(* IEC 61131-3 sources: SRCI_CLIENT_PLC/RobotLibrary/Library/POUs/General/MC_RobotTask, 1 file *)

(* ---- MC_RobotTaskFB.st ---- *)
/// Handles multiple mechanisms required for operation of the interface.
/// For maximal performance, this FB must be called after the function FB's,
/// so that the data can be written to the fieldbus in the same cycle as the start of FB occours
FUNCTION_BLOCK MC_RobotTaskFB EXTENDS RobotLibraryLogFB
// -------------------------------------------------------------------------
//  SRCI Robot Library
// -------------------------------------------------------------------------
//
//  Object:      RobotTaskFB
//  Author:      Thorsten Brach
//  Date:        2024-06-01
//
//  Description:
//
//
//  Copyright:
//    (C) 2024 Thorsten Brach. All rights reserved
//             Licensed under the MIT License.
//
//  Disclaimer:
//    This project is provided without any guarantee and can be used for
//    private and commercial purposes. Any use is at the user’s
//    own risk and responsibility.
//
// -------------------------------------------------------------------------
VAR_INPUT
  /// Set TRUE (default) to initialize the interface
  Enable            : BOOL;
  /// User defined robot name
  RobotName         : STRING(20);
  /// Current System Time
  SystemTime        : SystemTime;
  /// Online Change detected
  OnlineChange      : BOOL;
  /// Axes Group ID -> is used to uniquely identify each RA on a per RC basis.
  ///
  /// The IDs start with 0: an RC with only one RA uses ID 0.
  /// ST-FIX F138: spec V1.5.9 says 1 (one RA) and 1-15 (several RAs); this is an error of the spec
  /// (confirmed by PI), the SDK uses 0 too.
  AxesGroupID       : BYTE := 0;
  /// Configuration parameter
  ParCfg            : RobotTaskParCfg;
END_VAR

VAR_IN_OUT
  /// Inputs of PLC for communication from RC
  RobotInData       : ARRAY[*] OF BYTE;
  /// Outputs of PLC for communication to RC
  RobotOutData      : ARRAY[*] OF BYTE;
  ///  User data stored on the PLC according to Table 6-10
  UserData          : UserData;
  /// ToolData stored on PLC. For more information refer to 5.5.6.3
  ToolData          : ARRAY[*] OF Tool;
  /// LoadData stored on PLC.For more information refer to 5.5.6.4
  FrameData         : ARRAY[*] OF Frame;
  /// LoadData stored on PLC.For more information refer to 5.5.6.4
  LoadData          : ARRAY[*] OF Load;
  /// Work areas stored on PLC. For more information refer to 5.5.8
  WorkAreas         : ARRAY[*] OF RobotWorkArea;
  /// Software limits stored on PLC
  SWLimits          : SWLimits;
  /// Default dynamics stored on PLC. For more information refer to 5.5.7
  DefaultDynamics   : DefaultDynamics;
  /// Reference dynamics stored on PLC. For more information refer to 5.5.7
  ReferenceDynamics : ReferenceDynamics;
  /// System log on PLC
  SystemLog         : ARRAY[0..RobotLibraryParameter.SYSTEM_LOG_MAX ] OF STRING(RobotLibraryParameter.MESSAGE_TEXT_LEN);
  /// Message buffer on the PLC - For more information refer to 5.5.11
  MessageLog        : ARRAY[0..RobotLibraryParameter.MESSAGE_LOG_MAX] OF AlarmMessage;
  /// Robot assignment of function
  AxesGroup         : AxesGroup;
END_VAR

VAR_OUTPUT
  /// FB is being processed
  Busy              : BOOL;
  /// Interface is initialized (RI state: "Initialized").
  /// For more information on RI states refer to chapter 5.5.3.1.
  Initialized       : BOOL;
  /// Server and client were successfully synchronized (RI state: "Synchronized").
  /// For more information on the synchronization mechanism refer to chapter 5.6.7.
  Synchronized      : BOOL;
  /// An error occurred
  Error             : BOOL;
  /// ErrorID reported by RC for error identification according to Table 7-1
  ErrorID           : WORD;
  ErrorIdEnum       : RobotLibraryErrorIdEnum;
  ErrorAddTxt       : STRING(RobotLibraryConstants.MAX_ADD_TEXT_LENGTH);
  /// WarningID for warning identification reported during execution of command according to Table 7-3
  WarningID         : WORD;
  WarningIdEnum     : RobotLibraryWarningIdEnum;
  /// InfoID for info identification reported during execution of command according to Table 7-5
  InfoID            : WORD;
  InfoIdEnum        : RobotLibraryInfoIdEnum;
END_VAR

VAR
  /// internal copy of configuration parameter
 _parCfg                       : RobotTaskParCfg;

  /// internal ToolData for comparation to user ToolData
 _toolData                     : ARRAY[0..RobotLibraryParameter.TOOL_MAX       -1] OF Tool;
  /// internal FrameData for comparation to user FrameData
 _frameData                    : ARRAY[0..RobotLibraryParameter.FRAME_MAX      -1] OF Frame;
  /// internal LoadData for comparation to user LoadData
 _loadData                     : ARRAY[0..RobotLibraryParameter.LOAD_MAX       -1] OF Load;
  /// internal WorkAreas for comparation to user WorkAreas
 _workAreas                    : ARRAY[0..RobotLibraryParameter.WORK_AREAS_MAX -1] OF RobotWorkArea;
  /// internal Software limits for comparation to user Software limit
 _swLimits                     : SWLimits;
  /// internal default dynamics for comparation to user default dynamics
 _defaultDynamics              : DefaultDynamics;
  /// internal reference dynamics for comparation to user reference dynamics
 _referenceDynamics            : ReferenceDynamics;

  /// FB for exchange configuration
 _exchangeConfiguration        : MC_ExchangeConfigurationFB;
  /// FB for read robot data
 _readRobotData                : MC_ReadRobotDataFB;
  /// FB for read messaged
 _readMessages                 : MC_ReadMessagesFB;
  /// FB for read tool data
 _readToolData                 : MC_ReadToolDataFB;
  /// FB for read frame data
 _readFrameData                : MC_ReadFrameDataFB;
  /// FB for read load data
 _readLoadData                 : MC_ReadLoadDataFB;
  /// FB for read work area
 _readWorkArea                 : MC_ReadWorkAreaFB;
  /// FB for read robot software limits
 _readRobotSWLimits            : MC_ReadRobotSWLimitsFB;
  /// FB for read robot default dynamics
 _readRobotDefaultDynamics     : MC_ReadRobotDefaultDynamicsFB;
  /// FB for read robot reference dynamics
 _readRobotReferenceDynamics   : MC_ReadRobotReferenceDynamicsFB;

  /// FB for write tool data
 _writeToolData                : MC_WriteToolDataFB;
  /// FB for write frame data
 _writeFrameData               : MC_WriteFrameDataFB;
  /// FB for write load data
 _writeLoadData                : MC_WriteLoadDataFB;
  /// FB for write work area
 _writeWorkArea                : MC_WriteWorkAreaFB;
  /// FB for write robot software limits
 _writeRobotSWLimits           : MC_WriteRobotSWLimitsFB;
  /// FB for write robot default dynamics
 _writeRobotDefaultDynamics    : MC_WriteRobotDefaultDynamicsFB;
  /// FB for write robot reference dynamics
 _writeRobotReferenceDynamics  : MC_WriteRobotReferenceDynamicsFB;
  /// Send Buffer
  SendData                     : RobotLibrarySendDataFB;
  /// Recv Buffer
  RecvData                     : RobotLibraryRecvDataFB;
  /// Telegram
  Telegram                     : Telegram;

  /// internal step counter for command
 _stepCmd                      : DINT;
  /// internal timer for command
  {attribute 'hide'}
 _timerCmd                     : TON;
  /// internal timeout for command
  {attribute 'hide'}
 _timeoutCmd                   : TIME := T#5S;

  /// internal step counter for synchronisation of frame data
 _stepSyncFrameData            : DINT;
  /// internal timer for synchronisation of frame data
  {attribute 'hide'}
 _timerSyncFrameData           : TON;
  /// internal timeout for synchronisation of frame data
  {attribute 'hide'}
 _timeoutSyncFrameData         : TIME := T#5S;
   /// internal index for frame data synchronisation
 _syncIdxFrameData             : USINT;
  /// internal index for maximal amount of frames data( MIN(PLC,RC) )
 _syncIdxMaxFrameData          : DINT;

  /// internal step counter for synchronisation of load data
 _stepSyncLoadData             : DINT;
  /// internal timer for synchronisation of load data
  {attribute 'hide'}
 _timerSyncLoadData             : TON;
  /// internal timeout for synchronisation of load data
  {attribute 'hide'}
 _timeoutSyncLoadData           : TIME := T#5S;
  /// internal index for load data synchronisation
 _syncIdxLoadData               : USINT;
  /// internal index for maximal amount of load data ( MIN(PLC,RC) )
 _syncIdxMaxLoadData            : DINT;

  /// internal step counter for synchronisation of tool data
 _stepSyncToolData              : DINT;
  /// internal timer for synchronisation of tool data
  {attribute 'hide'}
 _timerSyncToolData             : TON;
  /// internal timeout for synchronisation of tool data
  {attribute 'hide'}
 _timeoutSyncToolData           : TIME := T#5S;
  /// internal index for tool data synchronisation
 _syncIdxToolData               : USINT;
  /// internal index for maximal amount of tool data ( MIN(PLC,RC) )
 _syncIdxMaxToolData            : DINT;

  /// internal step counter for synchronisation of work areas
 _stepSyncWorkArea            : DINT;
 /// internal timer for synchronisation of work areas
  {attribute 'hide'}
 _timerSyncWorkArea           : TON;
  /// internal timeout for synchronisation of work areas
  {attribute 'hide'}
 _timeoutSyncWorkArea         : TIME := T#5S;
  /// internal index for WorkArea synchronisation
 _syncIdxWorkArea             : USINT;
  /// internal index for maximal amount of Work Area( MIN(PLC,RC) )
 _syncIdxMaxWorkArea          : DINT;

  /// internal step counter for synchronisation of software limits
 _stepSyncSWLimits            : DINT;
  /// internal timer for synchronisation of software limits
  {attribute 'hide'}
 _timerSyncSWLimits           : TON;
  /// internal timeout for synchronisation of software limits
  {attribute 'hide'}
 _timeoutSyncSWLimits         : TIME := T#5S;

  /// internal step counter for synchronisation of default dynamics
 _stepSyncDefaultDynamics      : DINT;
  /// internal timer for synchronisation of default dynamics
  {attribute 'hide'}
 _timerSyncDefaultDynamics     : TON;
  /// internal timeout for synchronisation of default dynamics
  {attribute 'hide'}
 _timeoutSyncDefaultDynamics   : TIME := T#5S;

  /// internal step counter for synchronisation of reference dynamics
 _stepSyncReferenceDynamics    : DINT;
  /// internal timer for synchronisation of reference dynamics
  {attribute 'hide'}
 _timerSyncReferenceDynamics   : TON;
  /// internal timeout for synchronisation of reference dynamics
  {attribute 'hide'}
 _timeoutSyncReferenceDynamics : TIME := T#5S;

  /// Rising edge for enable
  {attribute 'hide'}
 _enable_R                    : R_TRIG;
  /// Falling edge for enable
  {attribute 'hide'}
 _enable_F                    : F_TRIG;

  /// Flag that indicated the the connection is alive (data exchange)
 _aliveBit                    : BOOL;
  /// last lifesign counter value
 _aliveValue                  : BYTE;
  /// timer for detecting alive state
 _aliveCheck                  : TON;
  /// rising edge for connection is alive
  {attribute 'hide'}
 _alive_R                     : R_TRIG;
  /// falling edge for connection is alive
  {attribute 'hide'}
 _alive_F                     : F_TRIG;
   /// last telegram state
 _lastTelegramState           : TelegramState   := TelegramState.UNDEFINED;
   /// last telegram control
 _lastTelegramControl         : ControlHalfByte := ControlHalfByte.NONE;
END_VAR

VAR // CONSTANT
  /// Lower array dimension of RobotInData
  ROBOT_IN_DATA_MIN   : DINT;
  /// Upper array dimension of RobotInData
  ROBOT_IN_DATA_MAX   : DINT;
  /// Size of RobotInData
  ROBOT_IN_DATA_SIZE  : UDINT;
  /// Lower array dimension of RobotOutData
  ROBOT_OUT_DATA_MIN  : DINT;
  /// Upper array dimension of RobotOutData
  ROBOT_OUT_DATA_MAX  : DINT;
  /// Size of RobotOutData
  ROBOT_OUT_DATA_SIZE : UDINT;
END_VAR

VAR CONSTANT
  {attribute 'hide'}
  FRAGMENT_HEADER_SIZE : UDINT := SIZEOF(TelegramPlcToRobFragmentHeader);
  /// Size of the comand header
  {attribute 'hide'}
  COMMAND_HEADER_SIZE  : UDINT := SIZEOF(TelegramPlcToRobCommandHeader);
  /// Size of the footer
  {attribute 'hide'}
  FOOTER_SIZE          : UDINT := 1;
  /// Minimal payload size for telegram
  {attribute 'hide'}
  MIN_PAYLOAD_SIZE     : UDINT := 1;
  /// Active command
  {attribute 'hide'}
  ACTIVE_CMD           : UDINT := 1;
  /// Buffered command
  {attribute 'hide'}
  BUFFER_CMD           : UDINT := 2;
  /// Empty command entry
  {attribute 'hide'}
  EMPTY_CMD_ENTRY      : AxesGroupAcyclicAcrEntryCmdBuffer := (State := BufferStateCmd.EMPTY);
  /// bitmask to mask the LifeSign out of the halfbyte
  {attribute 'hide'}
  LIFESIGN_BIT_MASK    : BYTE := 2#000_1111;
  /// Primary sequence
  {attribute 'hide'}
  PRIMARY_SEQUENCE     : DINT := 0;
  /// Secondary sequence
  {attribute 'hide'}
  SECONDARY_SEQUENCE   : DINT := 1;
  /// Empty Execution-Order-List entry
  {attribute 'hide'}
  EMPTY_EOL_ENTRY      : DINT := 0;
END_VAR

VAR
  /// ST-FIX F63: telegram sequence that is handled/filled first (lower Seq/Ack number)
  _seqSendFirst : DINT;
  /// ST-FIX F63: loop counter over the telegram sequences in Seq order
  _seqOrderIdx : DINT;
  /// ST-FIX F63: distance of two Seq numbers
  _seqDiff : DINT;
  /// ST-FIX F63: next Seq number
  _seqNext : UINT;
END_VAR

VAR
  /// ST-FIX F65: telegram sequence timeout (4 x LifeSignTimeOut without new Seq number)
  _seqAckTimeout : TON;
  /// ST-FIX F66: lifesign of header and footer differ -> frame is not processed
  _frameInvalid : BOOL;
  /// ST-FIX F79: last error state of the RC during the initialization (reported at the init timeout)
  _initErrorState : TelegramState;
END_VAR

VAR
  _turns : BYTE; // ST-FIX F60: turn number nibble
END_VAR

VAR
  _restartReset : BOOL; // ST-FIX F23: interface reset on the RC requested by a restart
END_VAR

VAR
  /// ST-FIX F132: identification of this instance (1..n, assigned in FB_init, kept by an online change)
 _instanceId : UDINT;
END_VAR

VAR_STAT
  /// ST-FIX F132: number of RobotTask instances created (source of _instanceId)
 _instanceCount   : UDINT;
  /// ST-FIX F132: instance that uses the telegram buffers of the entry (0 = free entry)
 _peripheryOwner  : ARRAY[1..PERIPHERY_ENTRIES] OF UDINT;
  /// ST-FIX F132: address of RobotInData of the entry
 _peripheryInAdr  : ARRAY[1..PERIPHERY_ENTRIES] OF PVOID;
  /// ST-FIX F132: address of RobotOutData of the entry
 _peripheryOutAdr : ARRAY[1..PERIPHERY_ENTRIES] OF PVOID;
END_VAR

VAR CONSTANT
  /// ST-FIX F132: number of RobotTask instances whose telegram buffers are checked
  PERIPHERY_ENTRIES : DINT := 16;
END_VAR

  // Get array dimension of RobotInData
  ROBOT_IN_DATA_MIN  := LOWER_BOUND  ( RobotInData,1);
  ROBOT_IN_DATA_MAX  := UPPER_BOUND  ( RobotInData,1);
  ROBOT_IN_DATA_SIZE := DINT_TO_UDINT( ROBOT_IN_DATA_MAX - ROBOT_IN_DATA_MIN + 1);

  // Get array dimension of RobotInData
  ROBOT_OUT_DATA_MIN  := LOWER_BOUND  ( RobotOutData,1);
  ROBOT_OUT_DATA_MAX  := UPPER_BOUND  ( RobotOutData,1);
  ROBOT_OUT_DATA_SIZE := DINT_TO_UDINT( ROBOT_OUT_DATA_MAX - ROBOT_OUT_DATA_MIN + 1);

  // ST-FIX F132: an AxesGroup and the telegram buffers belong to one RobotTask only (table 7-1:
  // 16#8007 / 16#8008); a second instance does nothing else, so it cannot disturb the first one
  IF ( NOT CheckAssignmentValid( AxesGroup    := AxesGroup,
                                 RobotInData  := RobotInData,
                                 RobotOutData := RobotOutData ) )
  THEN
    Error       := HasError;
    ErrorIdEnum := ErrorID;
    RETURN;
  END_IF

  HandleAxesGroup              ( AxesGroup         := AxesGroup,
  	                             ToolData          := ToolData,
  	                             FrameData         := FrameData,
  	                             LoadData          := LoadData,
  	                             WorkAreas         := WorkAreas,
  	                             SWLimits          := SWLimits,
  	                             DefaultDynamics   := DefaultDynamics,
  	                             ReferenceDynamics := ReferenceDynamics);

  HandleLifeSign               ( AxesGroup         := AxesGroup);
  HandleLogMessagesAck         ( AxesGroup         := AxesGroup);
  HandleInvalidFrames          ( AxesGroup         := AxesGroup, RobotInData := RobotInData);
  HandleTelegramStateCtrl      (                               );
  HandleAliveBit               ( RobotInData[1]                );
  HandleSeqAck                 ( AxesGroup         := AxesGroup);
  HandleUserData               ( AxesGroup         := AxesGroup, UserData := UserData );

  HandleSync                   ( AxesGroup         := AxesGroup,
                                 ToolData          := ToolData,
                                 FrameData         := FrameData,
                                 LoadData          := LoadData,
                                 WorkAreas         := WorkAreas,
                                 SWLimits          := SWLimits,
                                 DefaultDynamics   := DefaultDynamics,
                                 ReferenceDynamics := ReferenceDynamics);

  OnCall                       ( AxesGroup         := AxesGroup);
  OnExecRun                    ( AxesGroup         := AxesGroup);

  AxesGroupToTelegram          ( AxesGroup         := AxesGroup );

  CreateSendPayload            ( AxesGroup         := AxesGroup, RobotOutData := RobotOutData );
  IF ( NOT _frameInvalid ) // ST-FIX F66
  THEN
    ParseRecvPayload             ( AxesGroup         := AxesGroup, RobotInData  := RobotInData);
  END_IF

  AxesGroupFromTelegram        ( AxesGroup         := AxesGroup);

  // call internal functionblocks
  _exchangeConfiguration      ( Name := RobotName, ExecMode := ExecutionMode.PARALLEL, Priority := PriorityLevel.NORMAL, AxesGroup := AxesGroup );
  _readRobotData              ( Name := RobotName, ExecMode := ExecutionMode.PARALLEL, Priority := PriorityLevel.NORMAL, AxesGroup := AxesGroup );
  _readMessages               ( Name := RobotName, ExecMode := ExecutionMode.PARALLEL, Priority := PriorityLevel.NORMAL, AxesGroup := AxesGroup );
  _readToolData               ( UpdateSystemData := FALSE, // ST-FIX F16
   Name := RobotName, ExecMode := ExecutionMode.PARALLEL, Priority := PriorityLevel.NORMAL, AxesGroup := AxesGroup );
  _readFrameData              ( UpdateSystemData := FALSE, // ST-FIX F16
   Name := RobotName, ExecMode := ExecutionMode.PARALLEL, Priority := PriorityLevel.NORMAL, AxesGroup := AxesGroup );
  _readLoadData               ( UpdateSystemData := FALSE, // ST-FIX F16
   Name := RobotName, ExecMode := ExecutionMode.PARALLEL, Priority := PriorityLevel.NORMAL, AxesGroup := AxesGroup );
  _readWorkArea               ( UpdateSystemData := FALSE, // ST-FIX F16
   Name := RobotName, ExecMode := ExecutionMode.PARALLEL, Priority := PriorityLevel.NORMAL, AxesGroup := AxesGroup );
  _readRobotSWLimits          ( UpdateSystemData := FALSE, // ST-FIX F16
   Name := RobotName, ExecMode := ExecutionMode.PARALLEL, Priority := PriorityLevel.NORMAL, AxesGroup := AxesGroup );
  _readRobotDefaultDynamics   ( UpdateSystemData := FALSE, // ST-FIX F16
   Name := RobotName, ExecMode := ExecutionMode.PARALLEL, Priority := PriorityLevel.NORMAL, AxesGroup := AxesGroup );
  _readRobotReferenceDynamics ( UpdateSystemData := FALSE, // ST-FIX F16
   Name := RobotName, ExecMode := ExecutionMode.PARALLEL, Priority := PriorityLevel.NORMAL, AxesGroup := AxesGroup );
  _writeToolData              ( Name := RobotName, ExecMode := ExecutionMode.PARALLEL, Priority := PriorityLevel.NORMAL, AxesGroup := AxesGroup );
  _writeFrameData             ( Name := RobotName, ExecMode := ExecutionMode.PARALLEL, Priority := PriorityLevel.NORMAL, AxesGroup := AxesGroup );
  _writeLoadData              ( Name := RobotName, ExecMode := ExecutionMode.PARALLEL, Priority := PriorityLevel.NORMAL, AxesGroup := AxesGroup );
  _writeWorkArea              ( Name := RobotName, ExecMode := ExecutionMode.PARALLEL, Priority := PriorityLevel.NORMAL, AxesGroup := AxesGroup );
  _writeRobotSWLimits         ( Name := RobotName, ExecMode := ExecutionMode.PARALLEL, Priority := PriorityLevel.NORMAL, AxesGroup := AxesGroup );
  _writeRobotDefaultDynamics  ( Name := RobotName, ExecMode := ExecutionMode.PARALLEL, Priority := PriorityLevel.NORMAL, AxesGroup := AxesGroup );
  _writeRobotReferenceDynamics( Name := RobotName, ExecMode := ExecutionMode.PARALLEL, Priority := PriorityLevel.NORMAL, AxesGroup := AxesGroup );

  // Update SystemLog and MessageLog
  SystemLog  := AxesGroup.MessageLog.SystemLogs;
  MessageLog := AxesGroup.MessageLog.Messages;

END_FUNCTION_BLOCK

METHOD PRIVATE AxesGroupFromTelegram
VAR_IN_OUT
  /// Robot assignment of function
  AxesGroup    : AxesGroup;
END_VAR

  AxesGroupFromTelegramCyclic         (AxesGroup := AxesGroup);
  AxesGroupFromTelegramCyclicOptional (AxesGroup := AxesGroup);

END_METHOD

METHOD PRIVATE AxesGroupFromTelegramCyclic
VAR_IN_OUT
  /// Robot assignment of function
  AxesGroup : AxesGroup;
END_VAR

  // ---------------------------------
  // Mapp Telegramm to AxesGroup Data
  // ---------------------------------
  AxesGroup.Cyclic.RobToPlc.SRCIVersion    := Telegram.RobToPlc.Header.SRCIVersion ;
  AxesGroup.Cyclic.RobToPlc.LifeSign       := Telegram.RobToPlc.Header.LifeSign ;
  AxesGroup.Cyclic.RobToPlc.TelegramState  := Telegram.RobToPlc.Header.TelegramState ;
  AxesGroup.Cyclic.RobToPlc.StatusRobotArm := DwordToRaStatusWord(Telegram.RobToPlc.Header.StatusRobotArm);
  AxesGroup.Cyclic.RobToPlc.Override       := Telegram.RobToPlc.Header.Override ;

END_METHOD

METHOD PRIVATE AxesGroupFromTelegramCyclicOptional
VAR_IN_OUT
  /// Robot assignment of function
  AxesGroup: AxesGroup;
END_VAR

  // Sub ProgramData {{{
  AxesGroup.CyclicOptional.RobToPlc.SubProgramData.Data := Telegram.RobToPlc.CyclicOptional.SubProgramData.Data;
  // }}}

  // Cartesian position {{{
  AxesGroup.CyclicOptional.RobToPlc.CartesianPosition.Active                   :=                                     AxesGroup.CyclicOptional.RobToPlc.CartesianPosition.Active;
  AxesGroup.CyclicOptional.RobToPlc.CartesianPosition.X                        :=                                      Telegram.RobToPlc.CyclicOptional.CartesianPosition.X;
  AxesGroup.CyclicOptional.RobToPlc.CartesianPosition.Y                        :=                                      Telegram.RobToPlc.CyclicOptional.CartesianPosition.Y;
  AxesGroup.CyclicOptional.RobToPlc.CartesianPosition.Z                        :=                                      Telegram.RobToPlc.CyclicOptional.CartesianPosition.Z;
  AxesGroup.CyclicOptional.RobToPlc.CartesianPosition.Rx                       :=                                      Telegram.RobToPlc.CyclicOptional.CartesianPosition.Rx;
  AxesGroup.CyclicOptional.RobToPlc.CartesianPosition.Ry                       :=                                      Telegram.RobToPlc.CyclicOptional.CartesianPosition.Ry;
  AxesGroup.CyclicOptional.RobToPlc.CartesianPosition.Rz                       :=                                      Telegram.RobToPlc.CyclicOptional.CartesianPosition.Rz;
  AxesGroup.CyclicOptional.RobToPlc.CartesianPosition.Config.Shoulder          :=              WordToArmConfigShoulder(Telegram.RobToPlc.CyclicOptional.CartesianPosition.Config);
  AxesGroup.CyclicOptional.RobToPlc.CartesianPosition.Config.Elbow             :=              WordToArmConfigElbow   (Telegram.RobToPlc.CyclicOptional.CartesianPosition.Config);
  AxesGroup.CyclicOptional.RobToPlc.CartesianPosition.Config.Wrist             :=              WordToArmConfigWrist   (Telegram.RobToPlc.CyclicOptional.CartesianPosition.Config);
  _turns := GetHalfeByteLo(Telegram.RobToPlc.CyclicOptional.CartesianPosition.Turns_J2_J1); // ST-FIX F60: sign + magnitude (spec 5.5.4.4)
  AxesGroup.CyclicOptional.RobToPlc.CartesianPosition.TurnNumber.J1Turns := BYTE_TO_SINT(_turns AND 16#07);
  IF ( ( _turns AND 16#08 ) <> 0 )
  THEN
    AxesGroup.CyclicOptional.RobToPlc.CartesianPosition.TurnNumber.J1Turns := INT_TO_SINT(-SINT_TO_INT(AxesGroup.CyclicOptional.RobToPlc.CartesianPosition.TurnNumber.J1Turns));
  END_IF
  _turns := GetHalfeByteHi(Telegram.RobToPlc.CyclicOptional.CartesianPosition.Turns_J2_J1); // ST-FIX F60: sign + magnitude (spec 5.5.4.4)
  AxesGroup.CyclicOptional.RobToPlc.CartesianPosition.TurnNumber.J2Turns := BYTE_TO_SINT(_turns AND 16#07);
  IF ( ( _turns AND 16#08 ) <> 0 )
  THEN
    AxesGroup.CyclicOptional.RobToPlc.CartesianPosition.TurnNumber.J2Turns := INT_TO_SINT(-SINT_TO_INT(AxesGroup.CyclicOptional.RobToPlc.CartesianPosition.TurnNumber.J2Turns));
  END_IF
  _turns := GetHalfeByteLo(Telegram.RobToPlc.CyclicOptional.CartesianPosition.Turns_J4_J3); // ST-FIX F60: sign + magnitude (spec 5.5.4.4)
  AxesGroup.CyclicOptional.RobToPlc.CartesianPosition.TurnNumber.J3Turns := BYTE_TO_SINT(_turns AND 16#07);
  IF ( ( _turns AND 16#08 ) <> 0 )
  THEN
    AxesGroup.CyclicOptional.RobToPlc.CartesianPosition.TurnNumber.J3Turns := INT_TO_SINT(-SINT_TO_INT(AxesGroup.CyclicOptional.RobToPlc.CartesianPosition.TurnNumber.J3Turns));
  END_IF
  _turns := GetHalfeByteHi(Telegram.RobToPlc.CyclicOptional.CartesianPosition.Turns_J4_J3); // ST-FIX F60: sign + magnitude (spec 5.5.4.4)
  AxesGroup.CyclicOptional.RobToPlc.CartesianPosition.TurnNumber.J4Turns := BYTE_TO_SINT(_turns AND 16#07);
  IF ( ( _turns AND 16#08 ) <> 0 )
  THEN
    AxesGroup.CyclicOptional.RobToPlc.CartesianPosition.TurnNumber.J4Turns := INT_TO_SINT(-SINT_TO_INT(AxesGroup.CyclicOptional.RobToPlc.CartesianPosition.TurnNumber.J4Turns));
  END_IF
  _turns := GetHalfeByteLo(Telegram.RobToPlc.CyclicOptional.CartesianPosition.Turns_J6_J5); // ST-FIX F60: sign + magnitude (spec 5.5.4.4)
  AxesGroup.CyclicOptional.RobToPlc.CartesianPosition.TurnNumber.J5Turns := BYTE_TO_SINT(_turns AND 16#07);
  IF ( ( _turns AND 16#08 ) <> 0 )
  THEN
    AxesGroup.CyclicOptional.RobToPlc.CartesianPosition.TurnNumber.J5Turns := INT_TO_SINT(-SINT_TO_INT(AxesGroup.CyclicOptional.RobToPlc.CartesianPosition.TurnNumber.J5Turns));
  END_IF
  _turns := GetHalfeByteHi(Telegram.RobToPlc.CyclicOptional.CartesianPosition.Turns_J6_J5); // ST-FIX F60: sign + magnitude (spec 5.5.4.4)
  AxesGroup.CyclicOptional.RobToPlc.CartesianPosition.TurnNumber.J6Turns := BYTE_TO_SINT(_turns AND 16#07);
  IF ( ( _turns AND 16#08 ) <> 0 )
  THEN
    AxesGroup.CyclicOptional.RobToPlc.CartesianPosition.TurnNumber.J6Turns := INT_TO_SINT(-SINT_TO_INT(AxesGroup.CyclicOptional.RobToPlc.CartesianPosition.TurnNumber.J6Turns));
  END_IF
  AxesGroup.CyclicOptional.RobToPlc.CartesianPosition.TurnNumber.E1Turns := BYTE_TO_SINT(Telegram.RobToPlc.CyclicOptional.CartesianPosition.Turns_E1 AND 16#7F); // ST-FIX F60: sign + magnitude (spec 5.5.4.4)
  IF ( ( Telegram.RobToPlc.CyclicOptional.CartesianPosition.Turns_E1 AND 16#80 ) <> 0 )
  THEN
    AxesGroup.CyclicOptional.RobToPlc.CartesianPosition.TurnNumber.E1Turns := INT_TO_SINT(-SINT_TO_INT(AxesGroup.CyclicOptional.RobToPlc.CartesianPosition.TurnNumber.E1Turns));
  END_IF
  AxesGroup.CyclicOptional.RobToPlc.CartesianPosition.E1                       :=                                      Telegram.RobToPlc.CyclicOptional.CartesianPosition.E1;
  AxesGroup.CyclicOptional.RobToPlc.CartesianPosition.CoordinateSystem.ToolNo  :=                                      Telegram.RobToPlc.CyclicOptional.CartesianPosition.ToolNo; // ST-FIX F59: tool/frame of the returned position
  AxesGroup.CyclicOptional.RobToPlc.CartesianPosition.CurrentCoordinateSystem.ToolNo  :=                                      Telegram.RobToPlc.CyclicOptional.CartesianPosition.CurrentlyUsedToolNo;
  AxesGroup.CyclicOptional.RobToPlc.CartesianPosition.CoordinateSystem.FrameNo :=                                      Telegram.RobToPlc.CyclicOptional.CartesianPosition.FrameNo; // ST-FIX F59: tool/frame of the returned position
  AxesGroup.CyclicOptional.RobToPlc.CartesianPosition.CurrentCoordinateSystem.FrameNo :=                                      Telegram.RobToPlc.CyclicOptional.CartesianPosition.CurrentlyUsedFrameNo;
  // }}}

  // Joint position {{{
  AxesGroup.CyclicOptional.RobToPlc.JointPosition.Active := AxesGroup.CyclicOptional.RobToPlc.JointPosition.Active;
  AxesGroup.CyclicOptional.RobToPlc.JointPosition.J1     :=  Telegram.RobToPlc.CyclicOptional.JointPosition.J1;
  AxesGroup.CyclicOptional.RobToPlc.JointPosition.J2     :=  Telegram.RobToPlc.CyclicOptional.JointPosition.J2;
  AxesGroup.CyclicOptional.RobToPlc.JointPosition.J3     :=  Telegram.RobToPlc.CyclicOptional.JointPosition.J3;
  AxesGroup.CyclicOptional.RobToPlc.JointPosition.J4     :=  Telegram.RobToPlc.CyclicOptional.JointPosition.J4;
  AxesGroup.CyclicOptional.RobToPlc.JointPosition.J5     :=  Telegram.RobToPlc.CyclicOptional.JointPosition.J5;
  AxesGroup.CyclicOptional.RobToPlc.JointPosition.J6     :=  Telegram.RobToPlc.CyclicOptional.JointPosition.J6;
  AxesGroup.CyclicOptional.RobToPlc.JointPosition.E1     :=  Telegram.RobToPlc.CyclicOptional.JointPosition.E1;
  // }}}

  // Force {{{
  AxesGroup.CyclicOptional.RobToPlc.Force.Active          := AxesGroup.CyclicOptional.RobToPlc.Force.Active;
  AxesGroup.CyclicOptional.RobToPlc.Force.X               :=  Telegram.RobToPlc.CyclicOptional.Force.X;
  AxesGroup.CyclicOptional.RobToPlc.Force.Y               :=  Telegram.RobToPlc.CyclicOptional.Force.Y;
  AxesGroup.CyclicOptional.RobToPlc.Force.Z               :=  Telegram.RobToPlc.CyclicOptional.Force.Z;
  AxesGroup.CyclicOptional.RobToPlc.Force.Rx              :=  Telegram.RobToPlc.CyclicOptional.Force.Rx;
  AxesGroup.CyclicOptional.RobToPlc.Force.Ry              :=  Telegram.RobToPlc.CyclicOptional.Force.Ry;
  AxesGroup.CyclicOptional.RobToPlc.Force.Rz              :=  Telegram.RobToPlc.CyclicOptional.Force.Rz;
  // }}}

  // Current {{{
  AxesGroup.CyclicOptional.RobToPlc.Current.Active        := AxesGroup.CyclicOptional.RobToPlc.Current.Active;
  AxesGroup.CyclicOptional.RobToPlc.Current.J1            :=  Telegram.RobToPlc.CyclicOptional.Current.J1;
  AxesGroup.CyclicOptional.RobToPlc.Current.J2            :=  Telegram.RobToPlc.CyclicOptional.Current.J2;
  AxesGroup.CyclicOptional.RobToPlc.Current.J3            :=  Telegram.RobToPlc.CyclicOptional.Current.J3;
  AxesGroup.CyclicOptional.RobToPlc.Current.J4            :=  Telegram.RobToPlc.CyclicOptional.Current.J4;
  AxesGroup.CyclicOptional.RobToPlc.Current.J5            :=  Telegram.RobToPlc.CyclicOptional.Current.J5;
  AxesGroup.CyclicOptional.RobToPlc.Current.J6            :=  Telegram.RobToPlc.CyclicOptional.Current.J6;
  // }}}

  // Two Sequences {{{
  // }}}

  // Cartesian Position Extended
  AxesGroup.CyclicOptional.RobToPlc.CartesianPositionExt.Active := AxesGroup.CyclicOptional.RobToPlc.CartesianPositionExt.Active;
  AxesGroup.CyclicOptional.RobToPlc.CartesianPositionExt.E2     :=  Telegram.RobToPlc.CyclicOptional.CartesianPositionExt.E2;
  AxesGroup.CyclicOptional.RobToPlc.CartesianPositionExt.E3     :=  Telegram.RobToPlc.CyclicOptional.CartesianPositionExt.E3;
  AxesGroup.CyclicOptional.RobToPlc.CartesianPositionExt.E4     :=  Telegram.RobToPlc.CyclicOptional.CartesianPositionExt.E4;
  AxesGroup.CyclicOptional.RobToPlc.CartesianPositionExt.E5     :=  Telegram.RobToPlc.CyclicOptional.CartesianPositionExt.E5;
  AxesGroup.CyclicOptional.RobToPlc.CartesianPositionExt.E6     :=  Telegram.RobToPlc.CyclicOptional.CartesianPositionExt.E6;

  // Joint Position Extended
  AxesGroup.CyclicOptional.RobToPlc.JointPositionExt.Active     := AxesGroup.CyclicOptional.RobToPlc.JointPositionExt.Active;
  AxesGroup.CyclicOptional.RobToPlc.JointPositionExt.E2         :=  Telegram.RobToPlc.CyclicOptional.JointPositionExt.E2;
  AxesGroup.CyclicOptional.RobToPlc.JointPositionExt.E3         :=  Telegram.RobToPlc.CyclicOptional.JointPositionExt.E3;
  AxesGroup.CyclicOptional.RobToPlc.JointPositionExt.E4         :=  Telegram.RobToPlc.CyclicOptional.JointPositionExt.E4;
  AxesGroup.CyclicOptional.RobToPlc.JointPositionExt.E5         :=  Telegram.RobToPlc.CyclicOptional.JointPositionExt.E5;
  AxesGroup.CyclicOptional.RobToPlc.JointPositionExt.E6         :=  Telegram.RobToPlc.CyclicOptional.JointPositionExt.E6;

  // Force Extended
  AxesGroup.CyclicOptional.RobToPlc.ForceExt.Active             := AxesGroup.CyclicOptional.RobToPlc.ForceExt.Active;
  AxesGroup.CyclicOptional.RobToPlc.ForceExt.E1                 :=  Telegram.RobToPlc.CyclicOptional.ForceExt.E1;
  AxesGroup.CyclicOptional.RobToPlc.ForceExt.E2                 :=  Telegram.RobToPlc.CyclicOptional.ForceExt.E2;
  AxesGroup.CyclicOptional.RobToPlc.ForceExt.E3                 :=  Telegram.RobToPlc.CyclicOptional.ForceExt.E3;
  AxesGroup.CyclicOptional.RobToPlc.ForceExt.E4                 :=  Telegram.RobToPlc.CyclicOptional.ForceExt.E4;
  AxesGroup.CyclicOptional.RobToPlc.ForceExt.E5                 :=  Telegram.RobToPlc.CyclicOptional.ForceExt.E5;
  AxesGroup.CyclicOptional.RobToPlc.ForceExt.E6                 :=  Telegram.RobToPlc.CyclicOptional.ForceExt.E6;

  // Current Extended
  AxesGroup.CyclicOptional.RobToPlc.CurrentExt.Active           := AxesGroup.CyclicOptional.RobToPlc.CurrentExt.Active;
  AxesGroup.CyclicOptional.RobToPlc.CurrentExt.E1               :=  Telegram.RobToPlc.CyclicOptional.CurrentExt.E1;
  AxesGroup.CyclicOptional.RobToPlc.CurrentExt.E2               :=  Telegram.RobToPlc.CyclicOptional.CurrentExt.E2;
  AxesGroup.CyclicOptional.RobToPlc.CurrentExt.E3               :=  Telegram.RobToPlc.CyclicOptional.CurrentExt.E3;
  AxesGroup.CyclicOptional.RobToPlc.CurrentExt.E4               :=  Telegram.RobToPlc.CyclicOptional.CurrentExt.E4;
  AxesGroup.CyclicOptional.RobToPlc.CurrentExt.E5               :=  Telegram.RobToPlc.CyclicOptional.CurrentExt.E5;
  AxesGroup.CyclicOptional.RobToPlc.CurrentExt.E6               :=  Telegram.RobToPlc.CyclicOptional.CurrentExt.E6;

END_METHOD

METHOD PRIVATE AxesGroupToTelegram : DINT
VAR_IN_OUT
  /// Robot assignment of function
  AxesGroup : AxesGroup;
END_VAR

VAR
  /// internal index
 _idx                       : DINT;
  /// internal sequence index
 _seqIdx                    : DINT;
  /// internal fragment index
 _fragIdx                   : DINT;
  /// internal register index
 _regIdx                    : DINT;
  /// internal execution order list index
 _listIdx                   : DINT := 1;
  /// internal payload pointer
 _payLoadPtr                : DWORD;
  /// internal fragment action
 _fragmentAction            : FragmentAction;
  /// internal fragment action as string
 _fragmentActionString      : STRING;
  /// maximount amount of bytes per sequence
  SEQUENCE_MAX_PAYLOAD_SIZE : UDINT;
END_VAR

  // ST-FIX F63: the data of a telegram sequence is cleared in AxesGroupToTelegramSequence only
  // when it gets a new Seq number; a sequence that is not acknowledged yet is sent unchanged

  AxesGroupToTelegramHeader        (AxesGroup := AxesGroup);
  AxesGroupToTelegramCyclic        (AxesGroup := AxesGroup);
  AxesGroupToTelegramCyclicOptional(AxesGroup := AxesGroup);
  AxesGroupToTelegramSequence      (AxesGroup := AxesGroup);
  AxesGroupToTelegramFooter        (AxesGroup := AxesGroup);
  AxesGroupToTelegramLogging       (AxesGroup := AxesGroup);

END_METHOD

METHOD PRIVATE AxesGroupToTelegramCyclic : DINT
VAR_IN_OUT
  /// Robot assignment of function
  AxesGroup : AxesGroup;
END_VAR

  IF (AxesGroup.Cyclic.PlcToRob.ToolNo = -1 )
  THEN
    Telegram.PlcToRob.Cyclic.ToolNo  := 16#FF;
  ELSE
    Telegram.PlcToRob.Cyclic.ToolNo  := INT_TO_BYTE(AxesGroup.Cyclic.PlcToRob.ToolNo);
  END_IF

  IF (AxesGroup.Cyclic.PlcToRob.FrameNo = -1 )
  THEN
    Telegram.PlcToRob.Cyclic.FrameNo  := 16#FF;
  ELSE
    Telegram.PlcToRob.Cyclic.FrameNo  := INT_TO_BYTE(AxesGroup.Cyclic.PlcToRob.FrameNo);
  END_IF

END_METHOD

METHOD PRIVATE AxesGroupToTelegramCyclicOptional : DINT
VAR_IN_OUT
  /// Robot assignment of function
  AxesGroup : AxesGroup;
END_VAR

  // AxesGroup.CyclicOptional.PlcToRob.SubProgramData {{{
  IF (AxesGroup.CyclicOptional.PlcToRob.SubProgramData.Active)
  THEN
    Telegram.PlcToRob.CyclicOptional.SubProgramData.Data := AxesGroup.CyclicOptional.PlcToRob.SubProgramData.Data;
  END_IF
  // }}}

  // AxesGroup.CyclicOptional.PlcToRob.CartesianPosition  {{{
  IF (AxesGroup.CyclicOptional.PlcToRob.CartesianPosition.Active)
  THEN
    Telegram.PlcToRob.CyclicOptional.CartesianPosition.X           :=                  AxesGroup.CyclicOptional.PlcToRob.CartesianPosition.X;
    Telegram.PlcToRob.CyclicOptional.CartesianPosition.Y           :=                  AxesGroup.CyclicOptional.PlcToRob.CartesianPosition.Y;
    Telegram.PlcToRob.CyclicOptional.CartesianPosition.Z           :=                  AxesGroup.CyclicOptional.PlcToRob.CartesianPosition.Z;
    Telegram.PlcToRob.CyclicOptional.CartesianPosition.Rx          :=                  AxesGroup.CyclicOptional.PlcToRob.CartesianPosition.Rx;
    Telegram.PlcToRob.CyclicOptional.CartesianPosition.Ry          :=                  AxesGroup.CyclicOptional.PlcToRob.CartesianPosition.Ry;
    Telegram.PlcToRob.CyclicOptional.CartesianPosition.Rz          :=                  AxesGroup.CyclicOptional.PlcToRob.CartesianPosition.Rz;
    Telegram.PlcToRob.CyclicOptional.CartesianPosition.Turns_J2_J1 := CombineHalfSints(AxesGroup.CyclicOptional.PlcToRob.CartesianPosition.TurnNumber.J2Turns,
                                                                                       AxesGroup.CyclicOptional.PlcToRob.CartesianPosition.TurnNumber.J1Turns);
    Telegram.PlcToRob.CyclicOptional.CartesianPosition.Turns_J4_J3 := CombineHalfSints(AxesGroup.CyclicOptional.PlcToRob.CartesianPosition.TurnNumber.J4Turns,
                                                                                       AxesGroup.CyclicOptional.PlcToRob.CartesianPosition.TurnNumber.J3Turns);
    Telegram.PlcToRob.CyclicOptional.CartesianPosition.Turns_J6_J5 := CombineHalfSints(AxesGroup.CyclicOptional.PlcToRob.CartesianPosition.TurnNumber.J6Turns,
                                                                                       AxesGroup.CyclicOptional.PlcToRob.CartesianPosition.TurnNumber.J5Turns);
    // ST-FIX F60: sign + magnitude (spec 5.5.4.4)
    IF ( AxesGroup.CyclicOptional.PlcToRob.CartesianPosition.TurnNumber.E1Turns < 0 )
    THEN
      Telegram.PlcToRob.CyclicOptional.CartesianPosition.Turns_E1 := (INT_TO_BYTE(-SINT_TO_INT(AxesGroup.CyclicOptional.PlcToRob.CartesianPosition.TurnNumber.E1Turns)) AND 16#7F) OR 16#80;
    ELSE
      Telegram.PlcToRob.CyclicOptional.CartesianPosition.Turns_E1 := SINT_TO_BYTE(AxesGroup.CyclicOptional.PlcToRob.CartesianPosition.TurnNumber.E1Turns) AND 16#7F;
    END_IF
  END_IF
  // }}}

  // AxesGroup.CyclicOptional.PlcToRob.CartesianPositionExt {{{
  IF ( AxesGroup.CyclicOptional.PlcToRob.CartesianPositionExt.Active)
  THEN
    Telegram.PlcToRob.CyclicOptional.CartesianPositionExt.E2 := AxesGroup.CyclicOptional.PlcToRob.CartesianPositionExt.E2;
    Telegram.PlcToRob.CyclicOptional.CartesianPositionExt.E3 := AxesGroup.CyclicOptional.PlcToRob.CartesianPositionExt.E3;
    Telegram.PlcToRob.CyclicOptional.CartesianPositionExt.E4 := AxesGroup.CyclicOptional.PlcToRob.CartesianPositionExt.E4;
    Telegram.PlcToRob.CyclicOptional.CartesianPositionExt.E5 := AxesGroup.CyclicOptional.PlcToRob.CartesianPositionExt.E5;
    Telegram.PlcToRob.CyclicOptional.CartesianPositionExt.E6 := AxesGroup.CyclicOptional.PlcToRob.CartesianPositionExt.E6;
  END_IF
  // }}}

  // AxesGroup.CyclicOptional.PlcToRob.JointPosition {{{
  IF ( AxesGroup.CyclicOptional.PlcToRob.JointPosition.Active)
  THEN
    Telegram.PlcToRob.CyclicOptional.JointPosition.J1 := AxesGroup.CyclicOptional.PlcToRob.JointPosition.J1;
    Telegram.PlcToRob.CyclicOptional.JointPosition.J2 := AxesGroup.CyclicOptional.PlcToRob.JointPosition.J2;
    Telegram.PlcToRob.CyclicOptional.JointPosition.J3 := AxesGroup.CyclicOptional.PlcToRob.JointPosition.J3;
    Telegram.PlcToRob.CyclicOptional.JointPosition.J4 := AxesGroup.CyclicOptional.PlcToRob.JointPosition.J4;
    Telegram.PlcToRob.CyclicOptional.JointPosition.J5 := AxesGroup.CyclicOptional.PlcToRob.JointPosition.J5;
    Telegram.PlcToRob.CyclicOptional.JointPosition.J6 := AxesGroup.CyclicOptional.PlcToRob.JointPosition.J6;
    Telegram.PlcToRob.CyclicOptional.JointPosition.E1 := AxesGroup.CyclicOptional.PlcToRob.JointPosition.E1;
  END_IF
  // }}}

  // AxesGroup.CyclicOptional.PlcToRob.JointPositionExt {{{
  IF ( AxesGroup.CyclicOptional.PlcToRob.JointPositionExt.Active)
  THEN
    Telegram.PlcToRob.CyclicOptional.JointPositionExt.E2 := AxesGroup.CyclicOptional.PlcToRob.JointPositionExt.E2;
    Telegram.PlcToRob.CyclicOptional.JointPositionExt.E3 := AxesGroup.CyclicOptional.PlcToRob.JointPositionExt.E3;
    Telegram.PlcToRob.CyclicOptional.JointPositionExt.E4 := AxesGroup.CyclicOptional.PlcToRob.JointPositionExt.E4;
    Telegram.PlcToRob.CyclicOptional.JointPositionExt.E5 := AxesGroup.CyclicOptional.PlcToRob.JointPositionExt.E5;
    Telegram.PlcToRob.CyclicOptional.JointPositionExt.E6 := AxesGroup.CyclicOptional.PlcToRob.JointPositionExt.E6;
  END_IF
  // }}}

  // AxesGroup.CyclicOptional.PlcToRob.Force {{{
  IF ( AxesGroup.CyclicOptional.PlcToRob.Force.Active)
  THEN
    Telegram.PlcToRob.CyclicOptional.Force.X  := AxesGroup.CyclicOptional.PlcToRob.Force.X;
    Telegram.PlcToRob.CyclicOptional.Force.Y  := AxesGroup.CyclicOptional.PlcToRob.Force.Y;
    Telegram.PlcToRob.CyclicOptional.Force.Z  := AxesGroup.CyclicOptional.PlcToRob.Force.Z;
    Telegram.PlcToRob.CyclicOptional.Force.Rx := AxesGroup.CyclicOptional.PlcToRob.Force.Rx;
    Telegram.PlcToRob.CyclicOptional.Force.Ry := AxesGroup.CyclicOptional.PlcToRob.Force.Ry;
    Telegram.PlcToRob.CyclicOptional.Force.Rz := AxesGroup.CyclicOptional.PlcToRob.Force.Rz;
  END_IF
  // }}}

  // AxesGroup.CyclicOptional.PlcToRob.ForceExt {{{
  IF ( AxesGroup.CyclicOptional.PlcToRob.ForceExt.Active)
  THEN
    Telegram.PlcToRob.CyclicOptional.ForceExt.E1 := AxesGroup.CyclicOptional.PlcToRob.ForceExt.E1;
    Telegram.PlcToRob.CyclicOptional.ForceExt.E2 := AxesGroup.CyclicOptional.PlcToRob.ForceExt.E2;
    Telegram.PlcToRob.CyclicOptional.ForceExt.E3 := AxesGroup.CyclicOptional.PlcToRob.ForceExt.E3;
    Telegram.PlcToRob.CyclicOptional.ForceExt.E4 := AxesGroup.CyclicOptional.PlcToRob.ForceExt.E4;
    Telegram.PlcToRob.CyclicOptional.ForceExt.E5 := AxesGroup.CyclicOptional.PlcToRob.ForceExt.E5;
    Telegram.PlcToRob.CyclicOptional.ForceExt.E6 := AxesGroup.CyclicOptional.PlcToRob.ForceExt.E6;
  END_IF
  // }}}

END_METHOD

METHOD PRIVATE AxesGroupToTelegramFooter : DINT
VAR_IN_OUT
  /// Robot assignment of function
  AxesGroup : AxesGroup;
END_VAR

  Telegram.PlcToRob.Footer.LifeSign := GetHalfeByteLo(Telegram.PlcToRob.Header.FastStop_LifeSign);

END_METHOD

METHOD PRIVATE AxesGroupToTelegramHeader : DINT
VAR_IN_OUT
  /// Robot assignment of function
  AxesGroup : AxesGroup;
END_VAR

  Telegram.PlcToRob.Header.SRCIVersion               := VersionToByte(AxesGroup.Cyclic.PlcToRob.SRCIVersion);
  Telegram.PlcToRob.Header.FastStop_LifeSign         := CombineHalfBytes( HalfByteHi := AxesGroup.Cyclic.PlcToRob.FastStop, HalfByteLo := AxesGroup.Cyclic.PlcToRob.LifeSign );
  Telegram.PlcToRob.Header.TelegramLengthPlcToRob    := ParCfg.Com.TelegramLengthPlcToRob;
  Telegram.PlcToRob.Header.TelegramLengthRobToPlc    := ParCfg.Com.TelegramLengthRobToPlc;
  Telegram.PlcToRob.Header.AxesGroupID_Control       := CombineHalfBytes(HalfByteHi := AxesGroup.Cyclic.PlcToRob.AxesGroupID, HalfByteLo := AxesGroup.Cyclic.PlcToRob.Control);
  Telegram.PlcToRob.Header.Reserved                  := 0;
  Telegram.PlcToRob.Header.TelegramNumberPlcToRob    := PlcOptionalCyclicToUint(AxesGroup.Parameter.Plc.OptionalCyclic);
  Telegram.PlcToRob.Header.TelegramNumberRobToPlc    := RobOptionalCyclicToUint(AxesGroup.Parameter.Rob.OptionalCyclic);
  Telegram.PlcToRob.Header.ClientDate                := AxesGroup.Cyclic.PlcToRob.ClientDate;
  Telegram.PlcToRob.Header.ClientTime                := AxesGroup.Cyclic.PlcToRob.ClientTime;

END_METHOD

METHOD PRIVATE AxesGroupToTelegramLogging : DINT
VAR_IN_OUT
  /// Robot assignment of function
  AxesGroup : AxesGroup;
END_VAR

VAR
  /// internal sequence index
 _seqIdx                    : DINT;
  /// internal fragment index
 _fragIdx                   : DINT;
END_VAR

  FOR _seqIdx := 0 TO AxesGroup.State.SequenceCountSend
  DO
    // check new data ?
    IF ( AxesGroup.State.NewSEQ[_seqIdx] )
    THEN
      IF ( Telegram.PlcToRob.Sequence[_seqIdx].Header.PayloadLength > 0 )
      THEN
        // Create log entry
        CreateLogMessagePara4 ( Timestamp   := SystemTime,
                                MessageType := MessageType.CMD,
                                Severity    := Severity.DEBUG,
                                MessageCode := 0,
                                MessageText := 'SendData: SEQ = {1}, added Sequence [{2}] with PayloadLength = {3}, HeaderLength = {4}',
                                Para1       :=  UINT_TO_STRING(Telegram.PlcToRob.Sequence[_seqIdx].Header.SEQ_ACK),
                                Para2       :=  DINT_TO_STRING(_seqIdx),
                                Para3       :=  UINT_TO_STRING(Telegram.PlcToRob.Sequence[_seqIdx].Header.PayloadLength),
                                Para4       :=  DINT_TO_STRING(SIZEOF(Telegram.PlcToRob.Sequence[_seqIdx].Header)));
      END_IF

      FOR _fragIdx := 0 TO AxesGroup.State.FragmentCountSend[_seqIdx]
      DO
        IF ( Telegram.PlcToRob.Sequence[_seqIdx].Fragment[_fragIdx].Header.PayloadLength > 0 )
        THEN
          // Create log entry
          CreateLogMessagePara6 ( Timestamp   := SystemTime,
                                  MessageType := MessageType.CMD,
                                  Severity    := Severity.DEBUG,
                                  MessageCode := 0,
                                  MessageText := 'SendData: added Fragment [{1}] with PayloadLength = {2}, HeaderLength = {3}, CmdID <{4}>, Cmd <{5}> Fragment-Action Bits:{6}' ,
                                  Para1       := DINT_TO_STRING(_fragIdx),
                                  Para2       := UINT_TO_STRING            (Telegram.PlcToRob.Sequence[_seqIdx].Fragment[_fragIdx].Header.PayloadLength),
                                  Para3       := DINT_TO_STRING(SIZEOF     (Telegram.PlcToRob.Sequence[_seqIdx].Fragment[_fragIdx].Header)),
                                  Para4       := UINT_TO_STRING            (Telegram.PlcToRob.Sequence[_seqIdx].Fragment[_fragIdx].Header.CmdID),
                                  Para5       := CMD_TYPE_TO_STRING        (Telegram.PlcToRob.Sequence[_seqIdx].Fragment[_fragIdx].Command.Header.CmdType),
                                  Para6       := FRAGMENT_ACTION_TO_STRING (Telegram.PlcToRob.Sequence[_seqIdx].Fragment[_fragIdx].Header.FragmentAction));

          // Create log entry
          CreateLogMessagePara2 ( Timestamp   := SystemTime,
                                  MessageType := MessageType.CMD,
                                  Severity    := Severity.DEBUG,
                                  MessageCode := 0,
                                  MessageText := 'SendData: added Fragment [{1}] will be executed with ExecMode = [{2}]' ,
                                  Para1       := DINT_TO_STRING(_fragIdx),
                                  Para2       := EXECUTION_MODE_TO_STRING(Telegram.PlcToRob.Sequence[_seqIdx].Fragment[_fragIdx].Command.Header.ExecMode));

        END_IF
      END_FOR
    END_IF
  END_FOR

END_METHOD

METHOD PRIVATE AxesGroupToTelegramSequence : DINT
VAR_IN_OUT
  /// Robot assignment of function
  AxesGroup : AxesGroup;
END_VAR

VAR
  /// internal index
 _idx                       : DINT;
  /// internal sequence index
 _seqIdx                    : DINT;
   /// Amount of sequences
 _seqCount                  : DINT;

  /// internal fragment index
 _fragIdx                   : DINT;
  /// internal register index
 _regIdx                    : DINT;
  /// internal execution order list index
 _listIdx                   : DINT := 1;
  /// internal payload pointer
 _payLoadPtr                : DWORD;
  /// internal fragment action
 _fragmentAction            : FragmentAction;
  /// internal fragment action as string
 _fragmentActionString      : STRING;
  /// maximount amount of bytes per sequence
  SEQUENCE_MAX_PAYLOAD_SIZE : UDINT;

  /// current length of telegram
 _telegramLengthCurrent    : UINT;
END_VAR

  // Check 2nd sequence active ?
  // ST-FIX F67: remaining space for acyclic data at least 1 byte behind the sequence header
  IF ( CalculateSequencePayloadMax(AxesGroup := AxesGroup, Direction := ComDirection.PLC_TO_ROB,
                                   Sequence  := SequenceFlagEnum.PRIMARY_SEQUENCE) < 4 + 1 )
  THEN
    SetError( ErrorID := RobotLibraryErrorIdEnum.ERR_ACYCLIC_AREA_TO_SMALL_PLC_TO_ROB, Overwrite := FALSE );
    // Create log entry
    CreateLogMessage ( Timestamp   := SystemTime,
                       MessageType := MessageType.CMD,
                       Severity    := Severity.ERROR,
                       MessageCode := ErrorID,
                       MessageText := 'Telegram PLC -> RC: no space left for acyclic data');
    RETURN;
  END_IF
  IF ( CalculateSequencePayloadMax(AxesGroup := AxesGroup, Direction := ComDirection.ROB_TO_PLC,
                                   Sequence  := SequenceFlagEnum.PRIMARY_SEQUENCE) < 4 + 1 )
  THEN
    SetError( ErrorID := RobotLibraryErrorIdEnum.ERR_ACYCLIC_AREA_TO_SMALL_ROB_TO_PLC, Overwrite := FALSE );
    // Create log entry
    CreateLogMessage ( Timestamp   := SystemTime,
                       MessageType := MessageType.CMD,
                       Severity    := Severity.ERROR,
                       MessageCode := ErrorID,
                       MessageText := 'Telegram RC -> PLC: no space left for acyclic data');
    RETURN;
  END_IF

  IF ( _parCfg.Com.TwoSequences ) // ST-FIX F63: SEQUENCE_MAX_PAYLOAD_SIZE per sequence, see below
  THEN
    // inc sequence counter
   _seqCount := _seqCount + 1;
  END_IF

  FOR _seqOrderIdx := 0 TO _seqCount
  DO
    // ST-FIX F63: fill the sequence with the lower Seq number first (it is processed first)
    IF ( _seqOrderIdx = 0 )
    THEN
      _seqIdx := _seqSendFirst;
    ELSE
      _seqIdx := 1 - _seqSendFirst;
    END_IF
    // set current SEQ / ACk index
    Telegram.PlcToRob.Sequence[_seqIdx].Header.SEQ_ACK := AxesGroup.State.CurrentSEQ[_seqIdx];

    // only update telegram content if a new sequence SEQ is set
    IF ( AxesGroup.State.NewSEQ[_seqIdx] )
    THEN
      // only reset counters in case of new telegram to send
      // ST-FIX F63: each telegram sequence has its own data area (Fig. 5-205) and starts empty
      IF ( _seqIdx = PRIMARY_SEQUENCE )
      THEN
        SEQUENCE_MAX_PAYLOAD_SIZE := CalculateSequencePayloadMax(AxesGroup := AxesGroup,
                                                                 Direction := ComDirection.PLC_TO_ROB,
                                                                 Sequence  := SequenceFlagEnum.PRIMARY_SEQUENCE);
      ELSE
        SEQUENCE_MAX_PAYLOAD_SIZE := CalculateSequencePayloadMax(AxesGroup := AxesGroup,
                                                                 Direction := ComDirection.PLC_TO_ROB,
                                                                 Sequence  := SequenceFlagEnum.SECONDARY_SEQUENCE);
      END_IF
      Telegram.PlcToRob.Sequence[_seqIdx].Header.PayloadLength := 0;
      FOR _idx := 0 TO RobotLibraryParameter.FRAGMENT_MAX
      DO
        Telegram.PlcToRob.Sequence[_seqIdx].Fragment[_idx].Header.PayloadLength := 0;
      END_FOR
     _fragIdx := 0;
     _listIdx := 1;
      AxesGroup.State.FragmentCountSend[_seqIdx] := 0;

      // calc current telegram payload length
     _telegramLengthCurrent := 4 + Telegram.PlcToRob.Sequence[_seqIdx].Header.PayloadLength; // ST-FIX F63: sequence header + payload

      // Bedingung anpassen und TWO_SEQUENCES berücksichtigen
      WHILE ( _telegramLengthCurrent + FRAGMENT_HEADER_SIZE + MIN_PAYLOAD_SIZE <= SEQUENCE_MAX_PAYLOAD_SIZE ) // ST-FIX F63
      DO
        // Check command in Execution-Order-List available ?
        IF ( AxesGroup.Acyclic.ActiveCommandRegister.ExecutionOrderList[_listIdx] > EMPTY_EOL_ENTRY)
        THEN
          // set current SEQ / ACk index
          Telegram.PlcToRob.Sequence[_seqIdx].Header.SEQ_ACK := AxesGroup.State.CurrentSEQ[_seqIdx];

          // get active command register index
         _regIdx := AxesGroup.Acyclic.ActiveCommandRegister.ExecutionOrderList[_listIdx];

          // check State of the current ACR entry ?
          IF (( AxesGroup.Acyclic.ActiveCommandRegister.Register[_regIdx].Command[ACTIVE_CMD].State >= BufferStateCmd.CREATED  ) AND
              ( AxesGroup.Acyclic.ActiveCommandRegister.Register[_regIdx].Command[ACTIVE_CMD].State <= BufferStateCmd.SENDING  ))
          THEN
            // add size of fragement header
            Telegram.PlcToRob.Sequence[_seqIdx].Header.PayloadLength :=
              Telegram.PlcToRob.Sequence[_seqIdx].Header.PayloadLength + SIZEOF(Telegram.PlcToRob.Sequence[_seqIdx].Fragment[_fragIdx].Header);

            Telegram.PlcToRob.Sequence[_seqIdx].Fragment[_fragIdx].Header.CmdID          := AxesGroup.Acyclic.ActiveCommandRegister.Register[_regIdx].UniqueID;
            Telegram.PlcToRob.Sequence[_seqIdx].Fragment[_fragIdx].Header.Reserve        := 0;
            Telegram.PlcToRob.Sequence[_seqIdx].Fragment[_fragIdx].Header.FragmentAction := 0; // will be set below
            Telegram.PlcToRob.Sequence[_seqIdx].Fragment[_fragIdx].Header.PayloadPointer := AxesGroup.Acyclic.ActiveCommandRegister.Register[_regIdx].Command[ACTIVE_CMD].PayLoadPtr;

            // The 1st message resets the ACR entry on the server side
           _fragmentAction.Reset := (( AxesGroup.Acyclic.ActiveCommandRegister.Register[_regIdx].Command[ACTIVE_CMD].State      = BufferStateCmd.CREATED ) AND
                                     ( AxesGroup.Acyclic.ActiveCommandRegister.Register[_regIdx].Command[ACTIVE_CMD].PayLoadPtr = 0                      ));

            // Update messages must clear the ACR entry on the server side
           _fragmentAction.Clear := (( AxesGroup.Acyclic.ActiveCommandRegister.Register[_regIdx].Command[ACTIVE_CMD].State      = BufferStateCmd.UPDATE_AVAILABLE  ) AND
                                     ( AxesGroup.Acyclic.ActiveCommandRegister.Register[_regIdx].Command[ACTIVE_CMD].PayLoadPtr = 0                                ));

            // fill telegramm header - just for later debugging ( the header is part of the command payload itselfy ) {{{
            Telegram.PlcToRob.Sequence[_seqIdx].Fragment[_fragIdx].Command.Header.CmdType       := CombineBytesToUint ( AxesGroup.Acyclic.ActiveCommandRegister.Register[_regIdx].Command[ACTIVE_CMD].Payload[0],
                                                                                                                        AxesGroup.Acyclic.ActiveCommandRegister.Register[_regIdx].Command[ACTIVE_CMD].Payload[1]);
            Telegram.PlcToRob.Sequence[_seqIdx].Fragment[_fragIdx].Command.Header.ExecMode.0    :=                      AxesGroup.Acyclic.ActiveCommandRegister.Register[_regIdx].Command[ACTIVE_CMD].Payload[2].0;
            Telegram.PlcToRob.Sequence[_seqIdx].Fragment[_fragIdx].Command.Header.ExecMode.1    :=                      AxesGroup.Acyclic.ActiveCommandRegister.Register[_regIdx].Command[ACTIVE_CMD].Payload[2].1;
            Telegram.PlcToRob.Sequence[_seqIdx].Fragment[_fragIdx].Command.Header.ExecMode.2    :=                      AxesGroup.Acyclic.ActiveCommandRegister.Register[_regIdx].Command[ACTIVE_CMD].Payload[2].2;
            Telegram.PlcToRob.Sequence[_seqIdx].Fragment[_fragIdx].Command.Header.ExecMode.3    :=                      AxesGroup.Acyclic.ActiveCommandRegister.Register[_regIdx].Command[ACTIVE_CMD].Payload[2].3;
            Telegram.PlcToRob.Sequence[_seqIdx].Fragment[_fragIdx].Command.Header.Prio.0        :=                      AxesGroup.Acyclic.ActiveCommandRegister.Register[_regIdx].Command[ACTIVE_CMD].Payload[3].0;
            Telegram.PlcToRob.Sequence[_seqIdx].Fragment[_fragIdx].Command.Header.Prio.1        :=                      AxesGroup.Acyclic.ActiveCommandRegister.Register[_regIdx].Command[ACTIVE_CMD].Payload[3].1;
            Telegram.PlcToRob.Sequence[_seqIdx].Fragment[_fragIdx].Command.Header.Prio.2        :=                      AxesGroup.Acyclic.ActiveCommandRegister.Register[_regIdx].Command[ACTIVE_CMD].Payload[3].2;
            Telegram.PlcToRob.Sequence[_seqIdx].Fragment[_fragIdx].Command.Header.Prio.3        :=                      AxesGroup.Acyclic.ActiveCommandRegister.Register[_regIdx].Command[ACTIVE_CMD].Payload[3].3;
            Telegram.PlcToRob.Sequence[_seqIdx].Fragment[_fragIdx].Command.Header.ParSequence.0 :=                      AxesGroup.Acyclic.ActiveCommandRegister.Register[_regIdx].Command[ACTIVE_CMD].Payload[3].4;
            Telegram.PlcToRob.Sequence[_seqIdx].Fragment[_fragIdx].Command.Header.ParSequence.1 :=                      AxesGroup.Acyclic.ActiveCommandRegister.Register[_regIdx].Command[ACTIVE_CMD].Payload[3].5;
            Telegram.PlcToRob.Sequence[_seqIdx].Fragment[_fragIdx].Command.Header.ParSequence.2 :=                      AxesGroup.Acyclic.ActiveCommandRegister.Register[_regIdx].Command[ACTIVE_CMD].Payload[3].6;
            Telegram.PlcToRob.Sequence[_seqIdx].Fragment[_fragIdx].Command.Header.ParSequence.3 :=                      AxesGroup.Acyclic.ActiveCommandRegister.Register[_regIdx].Command[ACTIVE_CMD].Payload[3].7;
            // }}}
            // loop through the payload
            FOR _payLoadPtr := AxesGroup.Acyclic.ActiveCommandRegister.Register[_regIdx].Command[ACTIVE_CMD].PayLoadPtr TO AxesGroup.Acyclic.ActiveCommandRegister.Register[_regIdx].Command[ACTIVE_CMD].PayloadLen -1
            DO
              // copy payload
              Telegram.PlcToRob.Sequence[_seqIdx].Fragment[_fragIdx].Command.Payload[_payLoadPtr]
                := AxesGroup.Acyclic.ActiveCommandRegister.Register[_regIdx].Command[ACTIVE_CMD].Payload[_payLoadPtr];

              // inc current sequence payload length
              Telegram.PlcToRob.Sequence[_seqIdx].Header.PayloadLength
                := Telegram.PlcToRob.Sequence[_seqIdx].Header.PayloadLength + 1;

              // inc current fragment payload length
              Telegram.PlcToRob.Sequence[_seqIdx].Fragment[_fragIdx].Header.PayloadLength
                := Telegram.PlcToRob.Sequence[_seqIdx].Fragment[_fragIdx].Header.PayloadLength + 1;

              // inc payload pointer in active command register
              AxesGroup.Acyclic.ActiveCommandRegister.Register[_regIdx].Command[ACTIVE_CMD].PayLoadPtr
                := AxesGroup.Acyclic.ActiveCommandRegister.Register[_regIdx].Command[ACTIVE_CMD].PayLoadPtr + 1;

              // set command state
              IF ( AxesGroup.Acyclic.ActiveCommandRegister.Register[_regIdx].Command[ACTIVE_CMD].PayLoadPtr >= AxesGroup.Acyclic.ActiveCommandRegister.Register[_regIdx].Command[ACTIVE_CMD].PayLoadLen)
              THEN
                AxesGroup.Acyclic.ActiveCommandRegister.Register[_regIdx].Command[ACTIVE_CMD].State := BufferStateCmd.PROCESSED;
              ELSE
                AxesGroup.Acyclic.ActiveCommandRegister.Register[_regIdx].Command[ACTIVE_CMD].State := BufferStateCmd.SENDING;
              END_IF

              // calc current telegram payload length
             _telegramLengthCurrent := 4 + Telegram.PlcToRob.Sequence[_seqIdx].Header.PayloadLength; // ST-FIX F63: sequence header + payload

              // check limit reached ?
              IF ( _telegramLengthCurrent >= SEQUENCE_MAX_PAYLOAD_SIZE (* ST-FIX F63 *))
              THEN
                EXIT; // -> abort for loop
              END_IF
            END_FOR

            // check payload complete ?
           _fragmentAction.Complete := AxesGroup.Acyclic.ActiveCommandRegister.Register[_regIdx].Command[ACTIVE_CMD].PayLoadPtr
                                    >= AxesGroup.Acyclic.ActiveCommandRegister.Register[_regIdx].Command[ACTIVE_CMD].PayloadLen;

            // just for brakepoint
            IF (_fragmentAction.Complete)
            THEN
             _fragmentAction.Complete := _fragmentAction.Complete;
            END_IF

            // set fragment action
            Telegram.PlcToRob.Sequence[_seqIdx].Fragment[_fragIdx].Header.FragmentAction := FragmentActionToByte(_fragmentAction);
          END_IF
        END_IF

        // inc execution order list index
       _listIdx := _listIdx + 1;
        // inc fragment index
       _fragIdx := _fragIdx + 1;

        // check abort conditions
        IF (( _telegramLengthCurrent                                                >= SEQUENCE_MAX_PAYLOAD_SIZE (* ST-FIX F63 *)  ) OR  // Payload limit reached
            ( _fragIdx                                                              >=  RobotLibraryParameter.FRAGMENT_MAX ) OR  // Max fragment limit reached
            (  AxesGroup.Acyclic.ActiveCommandRegister.ExecutionOrderList[_listIdx]  =  EMPTY_EOL_ENTRY                    ))    // No entry in ExecutionOrderList left
        THEN
          EXIT;// -> Abort while loop
        END_IF
      END_WHILE

      AxesGroup.State.SequenceCountSend          := _seqCount; // ST-FIX F63
      AxesGroup.State.FragmentCountSend[_seqIdx] := _fragIdx;

    END_IF
  END_FOR

END_METHOD

METHOD CalculateCyclicDataLength : UINT
VAR_IN_OUT
  /// Robot assignment of function
  AxesGroup : AxesGroup;
END_VAR
VAR_INPUT
  /// Communication direction
  Direction : ComDirection;
END_VAR

VAR CONSTANT
  /// Size of the header
  ROB_TO_PLC_HEADER_SIZE : UINT := 10;
END_VAR

  // ------------------------------------
  // PLC -> ROB
  // ------------------------------------
  IF (Direction = ComDirection.PLC_TO_ROB)
  THEN
    // Add Header size
    CalculateCyclicDataLength := CalculateCyclicDataLength + SIZEOF(Telegram.PlcToRob.Header);
    // Add Cyclic size (ST-FIX F2: only with Cartesian Position RC -> PLC)
    IF ( AxesGroup.CyclicOptional.RobToPlc.CartesianPosition.Active )
    THEN
      CalculateCyclicDataLength := CalculateCyclicDataLength + SIZEOF(Telegram.PlcToRob.Cyclic);
    END_IF

    // Check SubProgramData active ?
    IF ( AxesGroup.CyclicOptional.PlcToRob.SubProgramData.Active )
    THEN
      // Add SubProgramData size
      CalculateCyclicDataLength := CalculateCyclicDataLength + SIZEOF(Telegram.PlcToRob.CyclicOptional.SubProgramData);
    END_IF

    // Check CartesianPosition active ?
    IF ( AxesGroup.CyclicOptional.PlcToRob.CartesianPosition.Active )
    THEN
      // Add CartesianPosition size
      CalculateCyclicDataLength := CalculateCyclicDataLength + SIZEOF(Telegram.PlcToRob.CyclicOptional.CartesianPosition);
    END_IF

    // Check JointPosition active ?
    IF ( AxesGroup.CyclicOptional.PlcToRob.JointPosition.Active )
    THEN
      // Add JointPosition size
      CalculateCyclicDataLength := CalculateCyclicDataLength + SIZEOF(Telegram.PlcToRob.CyclicOptional.JointPosition);
    END_IF

    // Check Force active ?
    IF ( AxesGroup.CyclicOptional.PlcToRob.Force.Active )
    THEN
      // Add Force size
      CalculateCyclicDataLength := CalculateCyclicDataLength + SIZEOF(Telegram.PlcToRob.CyclicOptional.Force);
    END_IF

    // Check CartesianPositionExt acive ?
    IF ( AxesGroup.CyclicOptional.PlcToRob.CartesianPositionExt.Active )
    THEN
      // Add CartesianPositionExt size
      CalculateCyclicDataLength := CalculateCyclicDataLength + SIZEOF(Telegram.PlcToRob.CyclicOptional.CartesianPositionExt);
    END_IF

    // Check JointPositionExt active ?
    IF ( AxesGroup.CyclicOptional.PlcToRob.JointPositionExt.Active )
    THEN
      // Add JointPositionExt size
      CalculateCyclicDataLength := CalculateCyclicDataLength + SIZEOF(Telegram.PlcToRob.CyclicOptional.JointPositionExt);
    END_IF

    // Check ForceExt active ?
    IF ( AxesGroup.CyclicOptional.PlcToRob.ForceExt.Active )
    THEN
      // Add ForceExt size
      CalculateCyclicDataLength := CalculateCyclicDataLength + SIZEOF(Telegram.PlcToRob.CyclicOptional.ForceExt);
    END_IF
  END_IF

  // ------------------------------------
  // ROB -> PLC
  // ------------------------------------
  IF (Direction = ComDirection.ROB_TO_PLC)
  THEN
    // Add Header size
    CalculateCyclicDataLength := CalculateCyclicDataLength + ROB_TO_PLC_HEADER_SIZE;
    // a constant, because SIZEOF(Telegram.RobToPlc.Header) counts the VersionStruct instead of one byte

    // Check SubProgramData active ?
    IF ( AxesGroup.CyclicOptional.RobToPlc.SubProgramData.Active )
    THEN
      // Add SubProgramData size
      CalculateCyclicDataLength := CalculateCyclicDataLength + SIZEOF(Telegram.RobToPlc.CyclicOptional.SubProgramData);
    END_IF

    // Check CartesianPosition active ?
    IF ( AxesGroup.CyclicOptional.RobToPlc.CartesianPosition.Active )
    THEN
      // Add CartesianPosition size
      CalculateCyclicDataLength := CalculateCyclicDataLength + SIZEOF(Telegram.RobToPlc.CyclicOptional.CartesianPosition);
    END_IF

    // Check JointPosition active ?
    IF ( AxesGroup.CyclicOptional.RobToPlc.JointPosition.Active )
    THEN
      // Add JointPosition size
      CalculateCyclicDataLength := CalculateCyclicDataLength + SIZEOF(Telegram.RobToPlc.CyclicOptional.JointPosition);
    END_IF

    // Check Force active ?
    IF ( AxesGroup.CyclicOptional.RobToPlc.Force.Active )
    THEN
      // Add Force size
      CalculateCyclicDataLength := CalculateCyclicDataLength + SIZEOF(Telegram.RobToPlc.CyclicOptional.Force);
    END_IF

    // Check Current acive ?
    IF ( AxesGroup.CyclicOptional.RobToPlc.Current.Active )
    THEN
      // Add Current size
      CalculateCyclicDataLength := CalculateCyclicDataLength + SIZEOF(Telegram.RobToPlc.CyclicOptional.Current);
    END_IF

    // Check CartesianPositionExt acive ?
    IF ( AxesGroup.CyclicOptional.RobToPlc.CartesianPositionExt.Active )
    THEN
      // Add CartesianPositionExt size
      CalculateCyclicDataLength := CalculateCyclicDataLength + SIZEOF(Telegram.RobToPlc.CyclicOptional.CartesianPositionExt);
    END_IF

    // Check JointPositionExt active ?
    IF ( AxesGroup.CyclicOptional.RobToPlc.JointPositionExt.Active )
    THEN
      // Add JointPositionExt size
      CalculateCyclicDataLength := CalculateCyclicDataLength + SIZEOF(Telegram.RobToPlc.CyclicOptional.JointPositionExt);
    END_IF

    // Check ForceExt active ?
    IF ( AxesGroup.CyclicOptional.RobToPlc.ForceExt.Active )
    THEN
      // Add ForceExt size
      CalculateCyclicDataLength := CalculateCyclicDataLength + SIZEOF(Telegram.RobToPlc.CyclicOptional.ForceExt);
    END_IF

    // Check CurrentExt active ?
    IF ( AxesGroup.CyclicOptional.RobToPlc.CurrentExt.Active )
    THEN
      // Add CurrentExt size
      CalculateCyclicDataLength := CalculateCyclicDataLength + SIZEOF(Telegram.RobToPlc.CyclicOptional.CurrentExt);
    END_IF
  END_IF

END_METHOD

METHOD CalculateSequencePayloadMax : UINT
VAR_IN_OUT
  /// Robot assignment of function
  AxesGroup : AxesGroup;
END_VAR
VAR_INPUT
  /// Communication direction
  Direction : ComDirection;
  /// Sequeunce
  Sequence : SequenceFlag;
END_VAR

VAR
  /// Length of the cyclic header
 _cyclicDataLength      : UINT;
  /// Acyclic area (ST-FIX F63)
 _area                  : UDINT;
END_VAR

  // calculate cyclic header length
  _cyclicDataLength := CalculateCyclicDataLength(AxesGroup := AxesGroup, Direction := Direction);

  // ST-FIX F63: acyclic area without the footer, halved for two sequences (spec Fig. 5-205)
  IF ( Direction = ComDirection.PLC_TO_ROB )
  THEN
    _area := UINT_TO_UDINT(_parCfg.Com.TelegramLengthPlcToRob) - UINT_TO_UDINT(_cyclicDataLength) - FOOTER_SIZE;
  ELSE
    _area := UINT_TO_UDINT(_parCfg.Com.TelegramLengthRobToPlc) - UINT_TO_UDINT(_cyclicDataLength) - FOOTER_SIZE;
  END_IF

  IF ( NOT _parCfg.Com.TwoSequences )
  THEN
    IF ( Sequence = SequenceFlag.PRIMARY_SEQUENCE )
    THEN
      CalculateSequencePayloadMax := UDINT_TO_UINT(_area);
    ELSE
      CalculateSequencePayloadMax := 0;
    END_IF
  ELSIF ( Sequence = SequenceFlag.PRIMARY_SEQUENCE )
  THEN
    CalculateSequencePayloadMax := UDINT_TO_UINT(_area / 2);
  ELSE
    CalculateSequencePayloadMax := UDINT_TO_UINT(_area - _area / 2);
  END_IF

END_METHOD

METHOD CalculateSequencePayloadStartAdr : UINT
VAR_IN_OUT
  /// Robot assignment of function
  AxesGroup : AxesGroup;
END_VAR
VAR_INPUT
  /// Communication direction
  Direction : ComDirection;
  /// Sequeunce
  Sequence : SequenceFlag;
END_VAR

VAR
  /// Length of the cyclic header
 _cyclicDataLength      : UINT;
  /// Length of the sequnce payload
 _sequencePayloadLength : UINT;
END_VAR

  // calculate cyclic header length
  _cyclicDataLength := CalculateCyclicDataLength(AxesGroup := AxesGroup, Direction := Direction);

  CASE (Sequence)
  OF

    SequenceFlag.PRIMARY_SEQUENCE   :

      // return start address
      CalculateSequencePayloadStartAdr := _cyclicDataLength;

    SequenceFlag.SECONDARY_SEQUENCE :

      // calculate sequence payload max
     _sequencePayloadLength
       := CalculateSequencePayloadMax( AxesGroup := AxesGroup,
                                       Direction := Direction,
                                       Sequence  := SequenceFlag.PRIMARY_SEQUENCE ); // ST-FIX F63: behind the area of the 1st sequence

      // return start address
      CalculateSequencePayloadStartAdr := _cyclicDataLength + _sequencePayloadLength;

  END_CASE

END_METHOD

METHOD PROTECTED CalculateTelegramLengthPlcToRob : UINT
VAR_IN_OUT
  /// Robot assignment of function
  AxesGroup : AxesGroup;
END_VAR
VAR
  /// length of the cyclic data block
 _cyclicDataLength : UINT;
END_VAR

  _cyclicDataLength := CalculateCyclicDataLength(AxesGroup := AxesGroup, Direction := ComDirection.PLC_TO_ROB);

  IF ( _parCfg.Com.TwoSequences )
  THEN
    CalculateTelegramLengthPlcToRob := _cyclicDataLength
                                      + SIZEOF(Telegram.PlcToRob.Sequence[  PRIMARY_SEQUENCE].Header)
                                      +       (Telegram.PlcToRob.Sequence[  PRIMARY_SEQUENCE].Header.PayloadLength)
                                      + SIZEOF(Telegram.PlcToRob.Sequence[SECONDARY_SEQUENCE].Header)
                                      +       (Telegram.PlcToRob.Sequence[SECONDARY_SEQUENCE].Header.PayloadLength)
                                      + SIZEOF(Telegram.PlcToRob.Footer);
  ELSE
    CalculateTelegramLengthPlcToRob := _cyclicDataLength
                                      + SIZEOF(Telegram.PlcToRob.Sequence[PRIMARY_SEQUENCE].Header)
                                      +       (Telegram.PlcToRob.Sequence[PRIMARY_SEQUENCE].Header.PayloadLength)
                                      + SIZEOF(Telegram.PlcToRob.Footer);
  END_IF

END_METHOD

/// ST-FIX F132: checks that the AxesGroup and the telegram buffers are not used by another RobotTask
/// (table 7-1: 16#8007 ERR_AXESGROUP_INVALID, 16#8008 ERR_PERIPHERY_INVALID) and registers them
METHOD PRIVATE CheckAssignmentValid : BOOL
VAR_IN_OUT
  /// Robot assignment of function
  AxesGroup    : AxesGroup;
  /// Inputs of PLC for communication from RC
  RobotInData  : ARRAY[*] OF BYTE;
  /// Outputs of PLC for communication to RC
  RobotOutData : ARRAY[*] OF BYTE;
END_VAR
VAR
  /// Loop index over the entries
 _idx     : DINT;
  /// Entry of this instance
 _own     : DINT;
  /// First free entry
 _free    : DINT;
  /// Address of RobotInData
 _inAdr   : PVOID;
  /// Address of RobotOutData
 _outAdr  : PVOID;
END_VAR

  CheckAssignmentValid := FALSE;

  // AxesGroup used by another RobotTask ?
  IF (( AxesGroup.State.RobotTaskId <> 0           ) AND
      ( AxesGroup.State.RobotTaskId <> _instanceId ))
  THEN
    IF ( ErrorID <> RobotLibraryErrorIdEnum.ERR_AXESGROUP_INVALID )
    THEN
      SetError( ErrorID := RobotLibraryErrorIdEnum.ERR_AXESGROUP_INVALID, Overwrite := TRUE );
      // Create log entry
      CreateLogMessagePara1 ( Timestamp   := SystemTime,
                              MessageType := MessageType.CMD,
                              Severity    := Severity.ERROR,
                              MessageCode := ErrorID,
                              MessageText := 'AxesGroup is already used by RobotTask {1}',
                              Para1       := UDINT_TO_STRING(AxesGroup.State.RobotTaskId));
    END_IF
    RETURN;
  END_IF

  // telegram buffers used by another RobotTask ?
  _inAdr  := ADR(RobotInData [ROBOT_IN_DATA_MIN ]);
  _outAdr := ADR(RobotOutData[ROBOT_OUT_DATA_MIN]);
  _own    := 0;
  _free   := 0;
  FOR _idx := 1 TO PERIPHERY_ENTRIES
  DO
    IF ( _peripheryOwner[_idx] = _instanceId )
    THEN
     _own := _idx;
    ELSIF ( _peripheryOwner[_idx] = 0 )
    THEN
      IF ( _free = 0 )
      THEN
       _free := _idx;
      END_IF
    ELSIF (( _peripheryInAdr [_idx] = _inAdr  ) OR
           ( _peripheryOutAdr[_idx] = _outAdr ))
    THEN
      IF ( ErrorID <> RobotLibraryErrorIdEnum.ERR_PERIPHERY_INVALID )
      THEN
        SetError( ErrorID := RobotLibraryErrorIdEnum.ERR_PERIPHERY_INVALID, Overwrite := TRUE );
        // Create log entry
        CreateLogMessagePara1 ( Timestamp   := SystemTime,
                                MessageType := MessageType.CMD,
                                Severity    := Severity.ERROR,
                                MessageCode := ErrorID,
                                MessageText := 'Telegram buffers are already used by RobotTask {1}',
                                Para1       := UDINT_TO_STRING(_peripheryOwner[_idx]));
      END_IF
      RETURN;
    END_IF
  END_FOR

  // register this instance (the addresses can change after an online change)
  IF ( _own = 0 )
  THEN
   _own := _free;
  END_IF
  IF ( _own > 0 )
  THEN
   _peripheryOwner [_own] := _instanceId;
   _peripheryInAdr [_own] := _inAdr;
   _peripheryOutAdr[_own] := _outAdr;
  END_IF
  AxesGroup.State.RobotTaskId := _instanceId;

  CheckAssignmentValid := TRUE;

END_METHOD

METHOD PROTECTED CheckParameterChanged : BOOL
VAR_IN_OUT
  /// Robot assignment of function
  AxesGroup    : AxesGroup;
END_VAR

VAR
  /// internal index for loops
 _idx : DINT;
END_VAR

  // Check initialization is already done ?
  IF ( NOT Initialized )
  THEN
    CheckParameterChanged := FALSE;
    RETURN;
  END_IF

  // compare memory
  CheckParameterChanged := ( SysDepMemCmp(pData1 := ADR(ParCfg), pData2 := ADR(_parCfg), DataLen := SIZEOF(ParCfg)) <> RobotLibraryConstants.OK );

  FOR _idx := SyncTime.DURING_START_UP TO SyncTime.AFTER_START_UP
  DO
    // Check Tool SyncMode changed ?
    IF ( _parCfg.Plc.Parameter.SynchronizationModes.Tool[_idx] <> ParCfg.Plc.Parameter.SynchronizationModes.Tool[_idx] )
    THEN
      // Set info
      SetInfo( InfoID := RobotLibraryInfoIdEnum.INFO_CHANGE_TOOL_SYNC_MODE_TO_NEGATIVE_ONLY_AT_PLC_START_ALLOWED, Overwrite := TRUE);

      // Create log entry
      CreateLogMessagePara3( Timestamp   := SystemTime,
                             MessageType := MessageType.CMD,
                             Severity    := Severity.INFO,
                             MessageCode := 0,
                             MessageText := 'SyncMode.Tool[{1}] changed from {2} to {3}, but this is only allowed at PLC start',
                             Para1       := SYNC_TIME_TO_STRING(_idx),
                             Para2       := SYNC_MODE_TO_STRING( ParCfg.Plc.Parameter.SynchronizationModes.Tool[_idx]),
                             Para3       := SYNC_MODE_TO_STRING(_parCfg.Plc.Parameter.SynchronizationModes.Tool[_idx]));
    END_IF

    // Check Frame SyncMode changed ?
    IF ( _parCfg.Plc.Parameter.SynchronizationModes.Frame[_idx] <> ParCfg.Plc.Parameter.SynchronizationModes.Frame[_idx] )
    THEN
      // Set info
      SetInfo( InfoID := RobotLibraryInfoIdEnum.INFO_CHANGE_FRAME_SYNC_MODE_TO_NEGATIVE_ONLY_AT_PLC_START_ALLOWED, Overwrite :=  TRUE);

      // Create log entry
      CreateLogMessagePara3( Timestamp   := SystemTime,
                             MessageType := MessageType.CMD,
                             Severity    := Severity.INFO,
                             MessageCode := 0,
                             MessageText := 'SyncMode.Frame[{1}] changed from {2} to {3}, but this is only allowed at PLC start',
                             Para1       := SYNC_TIME_TO_STRING(_idx),
                             Para2       := SYNC_MODE_TO_STRING( ParCfg.Plc.Parameter.SynchronizationModes.Frame[_idx]),
                             Para3       := SYNC_MODE_TO_STRING(_parCfg.Plc.Parameter.SynchronizationModes.Frame[_idx]));
    END_IF

    // Check Load SyncMode changed ?
    IF ( _parCfg.Plc.Parameter.SynchronizationModes.Load[_idx] <> ParCfg.Plc.Parameter.SynchronizationModes.Load[_idx] )
    THEN
      // Set info
      SetInfo( InfoID := RobotLibraryInfoIdEnum.INFO_CHANGE_LOAD_SYNC_MODE_TO_NEGATIVE_ONLY_AT_PLC_START_ALLOWED, Overwrite := TRUE);

      // Create log entry
      CreateLogMessagePara3( Timestamp   := SystemTime,
                             MessageType := MessageType.CMD,
                             Severity    := Severity.INFO,
                             MessageCode := 0,
                             MessageText := 'SyncMode.Load[{1}] changed from {2} to {3}, but this is only allowed at PLC start',
                             Para1       := SYNC_TIME_TO_STRING(_idx),
                             Para2       := SYNC_MODE_TO_STRING( ParCfg.Plc.Parameter.SynchronizationModes.Load[_idx]),
                             Para3       := SYNC_MODE_TO_STRING(_parCfg.Plc.Parameter.SynchronizationModes.Load[_idx]));
    END_IF

    // Check WorkAreas SyncMode changed ?
    IF ( _parCfg.Plc.Parameter.SynchronizationModes.WorkAreas[_idx] <> ParCfg.Plc.Parameter.SynchronizationModes.WorkAreas[_idx] )
    THEN
      // Set info
      SetInfo( InfoID := RobotLibraryInfoIdEnum.INFO_CHANGE_WORK_AREA_SYNC_MODE_TO_NEGATIVE_ONLY_AT_PLC_START_ALLOWED, Overwrite := TRUE);

      // Create log entry
      CreateLogMessagePara3( Timestamp   := SystemTime,
                             MessageType := MessageType.CMD,
                             Severity    := Severity.INFO,
                             MessageCode := 0,
                             MessageText := 'SyncMode.WorkAreas[{1}] changed from {2} to {3}, but this is only allowed at PLC start',
                             Para1       := SYNC_TIME_TO_STRING(_idx),
                             Para2       := SYNC_MODE_TO_STRING( ParCfg.Plc.Parameter.SynchronizationModes.WorkAreas[_idx]),
                             Para3       := SYNC_MODE_TO_STRING(_parCfg.Plc.Parameter.SynchronizationModes.WorkAreas[_idx]));
    END_IF

    // Check SWLimits SyncMode changed ?
    IF ( _parCfg.Plc.Parameter.SynchronizationModes.SWLimits[_idx] <> ParCfg.Plc.Parameter.SynchronizationModes.SWLimits[_idx] )
    THEN
      // Set info
      SetInfo( InfoID := RobotLibraryInfoIdEnum.INFO_CHANGE_SWLIMITS_SYNC_MODE_TO_NEGATIVE_ONLY_AT_PLC_START_ALLOWED, Overwrite := TRUE);

      // Create log entry
      CreateLogMessagePara3( Timestamp   := SystemTime,
                             MessageType := MessageType.CMD,
                             Severity    := Severity.INFO,
                             MessageCode := 0,
                             MessageText := 'SyncMode.SWLimits[{1}] changed from {2} to {3}, but this is only allowed at PLC start',
                             Para1       := SYNC_TIME_TO_STRING(_idx),
                             Para2       := SYNC_MODE_TO_STRING( ParCfg.Plc.Parameter.SynchronizationModes.SWLimits[_idx]),
                             Para3       := SYNC_MODE_TO_STRING(_parCfg.Plc.Parameter.SynchronizationModes.SWLimits[_idx]));
    END_IF

    // Check DefaultDynamics SyncMode changed ?
    IF ( _parCfg.Plc.Parameter.SynchronizationModes.DefaultDynamics[_idx] <> ParCfg.Plc.Parameter.SynchronizationModes.DefaultDynamics[_idx] )
    THEN
      // Set info
      SetInfo( InfoID := RobotLibraryInfoIdEnum.INFO_CHANGE_DEFAULT_DYNAMICS_SYNC_MODE_TO_NEGATIVE_ONLY_AT_PLC_START_ALLOWED, Overwrite := TRUE);

      // Create log entry
      CreateLogMessagePara3( Timestamp   := SystemTime,
                             MessageType := MessageType.CMD,
                             Severity    := Severity.INFO,
                             MessageCode := 0,
                             MessageText := 'SyncMode.DefaultDynamics[{1}] changed from {2} to {3}, but this is only allowed at PLC start',
                             Para1       := SYNC_TIME_TO_STRING(_idx),
                             Para2       := SYNC_MODE_TO_STRING( ParCfg.Plc.Parameter.SynchronizationModes.DefaultDynamics[_idx]),
                             Para3       := SYNC_MODE_TO_STRING(_parCfg.Plc.Parameter.SynchronizationModes.DefaultDynamics[_idx]));
    END_IF

    // Check ReferenceDynamics SyncMode changed ?
    IF ( _parCfg.Plc.Parameter.SynchronizationModes.ReferenceDynamics[_idx] <> ParCfg.Plc.Parameter.SynchronizationModes.ReferenceDynamics[_idx] )
    THEN
      // Set info
      SetInfo(InfoID := RobotLibraryInfoIdEnum.INFO_CHANGE_REFERENCE_DYNAMICS_SYNC_MODE_TO_NEGATIVE_ONLY_AT_PLC_START_ALLOWED, Overwrite := TRUE );

      // Create log entry
      CreateLogMessagePara3( Timestamp   := SystemTime,
                             MessageType := MessageType.CMD,
                             Severity    := Severity.INFO,
                             MessageCode := 0,
                             MessageText := 'SyncMode.ReferenceDynamics[{1}] changed from {2} to {3}, but this is only allowed at PLC start',
                             Para1       := SYNC_TIME_TO_STRING(_idx),
                             Para2       := SYNC_MODE_TO_STRING( ParCfg.Plc.Parameter.SynchronizationModes.ReferenceDynamics[_idx]),
                             Para3       := SYNC_MODE_TO_STRING(_parCfg.Plc.Parameter.SynchronizationModes.ReferenceDynamics[_idx]));
    END_IF

  END_FOR

  // Check Plc.OptionalCyclic changed ?
  IF ( PlcOptionalCyclicToUint(_parCfg.Plc.OptionalCyclic) <> PlcOptionalCyclicToUint(ParCfg.Plc.OptionalCyclic ))
  THEN
    // Set error
    SetWarning( WarningID := RobotLibraryWarningIdEnum.WARN_TELEGRAM_NO_CHANGED_DURING_OPERATION, Overwrite := TRUE ); // ST-FIX F68

    // Create log entry
    CreateLogMessagePara2( Timestamp   := SystemTime,
                           MessageType := MessageType.CMD,
                           Severity    := Severity.WARNING,
                           MessageCode := 0,
                           MessageText := 'ParCfg.Plc.OptionalCyclic changed after initialization from {1} to {2} -> Reinitialize by disabling and enabling the RobotTask',
                           Para1       := WORD_TO_STRING_BIN(PlcOptionalCyclicToUint(_parCfg.Plc.OptionalCyclic)),
                           Para2       := WORD_TO_STRING_BIN(PlcOptionalCyclicToUint( ParCfg.Plc.OptionalCyclic)));
  END_IF

  // Check Rob.OptionalCyclic changed ?
  IF ( RobOptionalCyclicToUint(_parCfg.Rob.OptionalCyclic) <> RobOptionalCyclicToUint(ParCfg.Rob.OptionalCyclic ))
  THEN
    // Set error
    SetWarning( WarningID := RobotLibraryWarningIdEnum.WARN_TELEGRAM_NO_CHANGED_DURING_OPERATION, Overwrite := TRUE ); // ST-FIX F68

    // Create log entry
    CreateLogMessagePara2( Timestamp   := SystemTime,
                           MessageType := MessageType.CMD,
                           Severity    := Severity.WARNING,
                           MessageCode := 0,
                           MessageText := 'ParCfg.Rob.OptionalCyclic changed after initialization from {1} to {2} -> Reinitialize by disabling and enabling the RobotTask',
                           Para1       := WORD_TO_STRING_BIN(RobOptionalCyclicToUint(_parCfg.Rob.OptionalCyclic)),
                           Para2       := WORD_TO_STRING_BIN(RobOptionalCyclicToUint( ParCfg.Rob.OptionalCyclic)));
  END_IF

END_METHOD

METHOD PROTECTED CheckParameterValid : BOOL
VAR_IN_OUT
  /// Robot assignment of function
  AxesGroup : AxesGroup;
END_VAR

  // init return value
  CheckParameterValid := TRUE;

  // Check ParCfg.Com.TelegramLengthPlcToRob
  IF ( ParCfg.Com.TelegramLengthPlcToRob < 128 )
  THEN
    // Set Warning
    SetWarning( WarningID := RobotLibraryWarningIdEnum.WARN_ACYCLIC_RANGE_PLC_TO_ROB_VERY_SMALL, Overwrite := TRUE );
  END_IF

  // Check ParCfg.Com.TelegramLengthRobToPlc
  IF ( ParCfg.Com.TelegramLengthRobToPlc < 128 )
  THEN
    // Set Warning
    SetWarning( WarningID := RobotLibraryWarningIdEnum.WARN_ACYCLIC_RANGE_ROB_TO_PLC_VERY_SMALL, Overwrite := TRUE );
  END_IF

  // Region ParCfg.Com {{{

  // Check LifeSignTimeout
  IF ( ParCfg.Com.LifeSignTimeOut < T#10MS )
  THEN
    // set to valid min value
    ParCfg.Com.LifeSignTimeOut := T#10MS;

    // Set info
    SetInfo( InfoID := RobotLibraryInfoIdEnum.INFO_LIFESIGN_TIMEOUT_TO_SMALL_AND_SET_TO_10MS, Overwrite := TRUE);

    // Create log entry
    CreateLogMessagePara1 ( Timestamp   := SystemTime,
                            MessageType := MessageType.CMD,
                            Severity    := Severity.INFO,
                            MessageCode := 0,
                            MessageText := 'LifeSignTimeout to small and set from {1}ms to 10ms',
                            Para1       := TIME_TO_STRING(ParCfg.Com.LifeSignTimeOut));
  END_IF

  // Check ParCfg.Com.TelegramLengthPlcToRob
  IF (( ParCfg.Com.TelegramLengthPlcToRob < 64                  ) OR
      ( ParCfg.Com.TelegramLengthPlcToRob > ROBOT_OUT_DATA_SIZE ))
  THEN
    // parameter(s) not valid
    CheckParameterValid := FALSE;

    // Set error
    SetError( ErrorID := RobotLibraryErrorIdEnum.ERR_TELEGRAM_LENGTH_MISMATCH_0x80A3, Overwrite := TRUE );

    // Create log entry
    CreateLogMessagePara1 ( Timestamp   := SystemTime,
                            MessageType := MessageType.CMD,
                            Severity    := Severity.INFO,
                            MessageCode := 0,
                            MessageText :=               'ParCfg.Com.TelegramLengthPlcToRob {1} invalid',
                            Para1       := UINT_TO_STRING(ParCfg.Com.TelegramLengthPlcToRob));
    // no further validation
    RETURN;
  END_IF

  // Check ParCfg.Com.TelegramLengthRobToPlc
  IF (( ParCfg.Com.TelegramLengthRobToPlc < 64                 ) OR
      ( ParCfg.Com.TelegramLengthRobToPlc > ROBOT_IN_DATA_SIZE ))
  THEN
    // parameter(s) not valid
    CheckParameterValid := FALSE;

    // Set error
    SetError( ErrorID := RobotLibraryErrorIdEnum.ERR_TELEGRAM_LENGTH_MISMATCH_0x80A3, Overwrite := TRUE );

    // Create log entry
    CreateLogMessagePara1 ( Timestamp   := SystemTime,
                            MessageType := MessageType.CMD,
                            Severity    := Severity.INFO,
                            MessageCode := 0,
                            MessageText :=               'ParCfg.Com.TelegramLengthRobToPlc {1} invalid',
                            Para1       := UINT_TO_STRING(ParCfg.Com.TelegramLengthRobToPlc));
    // no further validation
    RETURN;
  END_IF
  // ST-FIX F63: two telegram sequences must be activated in both directions and for the layout
  IF ( ParCfg.Plc.OptionalCyclic.UseTwoSequences <> ParCfg.Rob.OptionalCyclic.UseTwoSequences ) OR
     ( ParCfg.Plc.OptionalCyclic.UseTwoSequences <> ParCfg.Com.TwoSequences                  )
  THEN
    CheckParameterValid := FALSE;
    SetError( ErrorID := RobotLibraryErrorIdEnum.ERR_TELEGRAM_NUMBER_INVALID_0x80AB, Overwrite := TRUE );
    CreateLogMessage( Timestamp   := SystemTime,
                      MessageType := MessageType.CMD,
                      Severity    := Severity.ERROR,
                      MessageCode := 0,
                      MessageText := 'TwoSequences must be set in Com and in Plc/Rob.OptionalCyclic');
    RETURN;
  END_IF
  // EndRegion }}}

  // Region ParCfg.Rob.OptionalCyclic {{{

  // Check configuration if optional cyclic CartesianPosition valid ?
  // ST-FIX F137: the extended cartesian position cannot be used without the cartesian position ->
  // the cartesian position is activated automatically (spec 6.4.2 and InfoID 16#6002, table 7-6);
  // before: both together were rejected and the extended position was switched off
  IF ( ParCfg.Rob.OptionalCyclic.UseCartesianPositionExt AND NOT ParCfg.Rob.OptionalCyclic.UseCartesianPosition )
  THEN
    // set to valid configuration
    ParCfg.Rob.OptionalCyclic.UseCartesianPosition    := TRUE;

    // Set info
    SetInfo( InfoID := RobotLibraryInfoIdEnum.INFO_RECV_EXT_CART_POS_NOT_USABLE_WITH_RECV_CART_POS, Overwrite := TRUE);

    // Create log entry
    CreateLogMessage( Timestamp   := SystemTime,
                      MessageType := MessageType.CMD,
                      Severity    := Severity.INFO,
                      MessageCode := 0,
                      MessageText := 'UseCartesianPositionExt cannot be used without UseCartesianPosition -> UseCartesianPosition is automatically activated');
  END_IF

  // Check configuration if optional cyclic JointPosition valid ?
  // ST-FIX F137: the extended joint position cannot be used without the joint position -> the joint
  // position is activated automatically (spec 6.4.2 and InfoID 16#6003, table 7-6); before: the check
  // (both together rejected) was switched off with AND FALSE
  IF ( ParCfg.Rob.OptionalCyclic.UseJointPositionExt AND NOT ParCfg.Rob.OptionalCyclic.UseJointPosition )
  THEN
    // set to valid configuration
    ParCfg.Rob.OptionalCyclic.UseJointPosition    := TRUE;

    // Set info
    SetInfo( InfoID := RobotLibraryInfoIdEnum.INFO_RECV_EXT_JOINT_POS_NOT_USABLE_WITH_RECV_JOINT_POS, Overwrite := TRUE);

    // Create log entry
    CreateLogMessage( Timestamp   := SystemTime,
                      MessageType := MessageType.CMD,
                      Severity    := Severity.INFO,
                      MessageCode := 0,
                      MessageText := 'UseJointPositionExt cannot be used without UseJointPosition -> UseJointPosition is automatically activated');
  END_IF
  // EndRegion }}}

  // Region ParCfg.Parameter.SynchronizationModes {{{

  // Check ToolData synchronisation mode during startup
  IF (( ParCfg.Plc.Parameter.SynchronizationModes.Tool[SyncTime.DURING_START_UP] <  SyncMode.NO_SYNCHRONIZATION ) OR
      ( ParCfg.Plc.Parameter.SynchronizationModes.Tool[SyncTime.DURING_START_UP] >= SyncMode.AUTOMATIC          )) // Automatic is not allowed during startup
  THEN
    // ST-FIX F130: only the warning of the data set (spec: no error); the RobotTask is initialized,
    // the data set is not synchronized (SyncModesValid in the HandleSync... methods)
    SetWarning( WarningID := RobotLibraryWarningIdEnum.WARN_TOOL_DATA_SYNC_MODE_INVALID, Overwrite := TRUE );

    // Create log entry
    CreateLogMessagePara1 ( Timestamp   := SystemTime,
                            MessageType := MessageType.CMD,
                            Severity    := Severity.INFO,
                            MessageCode := 0,
                            MessageText :=                    'ParCfg.Plc.Parameter.SynchronizationModes.Tool[SyncTime.DURING_START_UP] invalid SyncMode {1}',
                            Para1       := SYNC_MODE_TO_STRING(ParCfg.Plc.Parameter.SynchronizationModes.Tool[SyncTime.DURING_START_UP]));
  END_IF

  // Check ToolData synchronisation mode after startup
  IF (( ParCfg.Plc.Parameter.SynchronizationModes.Tool[SyncTime.AFTER_START_UP] < SyncMode.NO_SYNCHRONIZATION ) OR
      ( ParCfg.Plc.Parameter.SynchronizationModes.Tool[SyncTime.AFTER_START_UP] > SyncMode.AUTOMATIC          ))
  THEN
    // ST-FIX F130: only the warning of the data set (spec: no error); the RobotTask is initialized,
    // the data set is not synchronized (SyncModesValid in the HandleSync... methods)
    SetWarning( WarningID := RobotLibraryWarningIdEnum.WARN_TOOL_DATA_SYNC_MODE_INVALID, Overwrite := TRUE);

    // Create log entry
    CreateLogMessagePara1 ( Timestamp   := SystemTime,
                            MessageType := MessageType.CMD,
                            Severity    := Severity.INFO,
                            MessageCode := 0,
                            MessageText :=                    'ParCfg.Plc.Parameter.SynchronizationModes.Tool[SyncTime.AFTER_START_UP] invalid SyncMode {1}',
                            Para1       := SYNC_MODE_TO_STRING(ParCfg.Plc.Parameter.SynchronizationModes.Tool[SyncTime.AFTER_START_UP]));
  END_IF

  // Check FrameData synchronisation mode during startup
  IF (( ParCfg.Plc.Parameter.SynchronizationModes.Frame[SyncTime.DURING_START_UP] <  SyncMode.NO_SYNCHRONIZATION ) OR
      ( ParCfg.Plc.Parameter.SynchronizationModes.Frame[SyncTime.DURING_START_UP] >= SyncMode.AUTOMATIC          )) // Automatic is not allowed during startup
  THEN
    // ST-FIX F130: only the warning of the data set (spec: no error); the RobotTask is initialized,
    // the data set is not synchronized (SyncModesValid in the HandleSync... methods)
    SetWarning( WarningID := RobotLibraryWarningIdEnum.WARN_FRAME_DATA_SYNC_MODE_INVALID, Overwrite := FALSE);

    // Create log entry
    CreateLogMessagePara1 ( Timestamp   := SystemTime,
                            MessageType := MessageType.CMD,
                            Severity    := Severity.INFO,
                            MessageCode := 0,
                            MessageText :=                    'ParCfg.Plc.Parameter.SynchronizationModes.Frame[SyncTime.DURING_START_UP] invalid SyncMode {1}',
                            Para1       := SYNC_MODE_TO_STRING(ParCfg.Plc.Parameter.SynchronizationModes.Frame[SyncTime.DURING_START_UP]));
  END_IF

  // Check FrameData synchronisation mode after startup
  IF (( ParCfg.Plc.Parameter.SynchronizationModes.Frame[SyncTime.AFTER_START_UP] < SyncMode.NO_SYNCHRONIZATION ) OR
      ( ParCfg.Plc.Parameter.SynchronizationModes.Frame[SyncTime.AFTER_START_UP] > SyncMode.AUTOMATIC          ))
  THEN
    // ST-FIX F130: only the warning of the data set (spec: no error); the RobotTask is initialized,
    // the data set is not synchronized (SyncModesValid in the HandleSync... methods)
    SetWarning( WarningID := RobotLibraryWarningIdEnum.WARN_FRAME_DATA_SYNC_MODE_INVALID, Overwrite := TRUE);

    // Create log entry
    CreateLogMessagePara1 ( Timestamp   := SystemTime,
                            MessageType := MessageType.CMD,
                            Severity    := Severity.INFO,
                            MessageCode := 0,
                            MessageText :=                    'ParCfg.Plc.Parameter.SynchronizationModes.Frame[SyncTime.AFTER_START_UP] invalid SyncMode {1}',
                            Para1       := SYNC_MODE_TO_STRING(ParCfg.Plc.Parameter.SynchronizationModes.Frame[SyncTime.AFTER_START_UP]));
  END_IF

  // Check LoadData synchronisation mode during startup
  IF (( ParCfg.Plc.Parameter.SynchronizationModes.Load[SyncTime.DURING_START_UP] <  SyncMode.NO_SYNCHRONIZATION ) OR
      ( ParCfg.Plc.Parameter.SynchronizationModes.Load[SyncTime.DURING_START_UP] >= SyncMode.AUTOMATIC          )) // Automatic is not allowed during startup
  THEN
    // ST-FIX F130: only the warning of the data set (spec: no error); the RobotTask is initialized,
    // the data set is not synchronized (SyncModesValid in the HandleSync... methods)
    SetWarning ( WarningID := RobotLibraryWarningIdEnum.WARN_LOAD_DATA_SYNC_MODE_INVALID, Overwrite := TRUE);
